   729: '-YB4 OP3_RESERVE_1', class Errors, trigger "DB_ALARM_OP3_M_3" bit 8
   730: '-YB4 OP3_RESERVE_2', class Errors, trigger "DB_ALARM_OP3_M_3" bit 9
   731: '-YB4 OP3_RESERVE_3', class Errors, trigger "DB_ALARM_OP3_M_3" bit 10
   732: '-YB4 OP3_RESERVE_4', class Errors, trigger "DB_ALARM_OP3_M_3" bit 11
   733: '-YB4 OP3_RESERVE_5', class Errors, trigger "DB_ALARM_OP3_M_3" bit 12
   734: '-YB4 OP3_RESERVE_6', class Errors, trigger "DB_ALARM_OP3_M_3" bit 13
   735: '-YB4 OP3_RESERVE_7', class Errors, trigger "DB_ALARM_OP3_M_3" bit 14
   736: '-YB4 OP3_RESERVE_8', class Errors, trigger "DB_ALARM_OP3_M_3" bit 15
   737: 'OP3_N0 -YB5 Nespecifikovaný režim motoru AUTOMAT/MANUAL', class Errors, trigger "DB_ALARM_OP3_M_4" bit 0
   738: 'OP3_N0 -YB5 Externí alarm err 1', class Errors, trigger "DB_ALARM_OP3_M_4" bit 1
   739: 'OP3_N0 -YB5 Externí alarm err 2', class Errors, trigger "DB_ALARM_OP3_M_4" bit 2
   740: 'OP3_N0 -YB5 Externí alarm err 3', class Errors, trigger "DB_ALARM_OP3_M_4" bit 3
   741: 'OP3_N0 -YB5 Motor nemá splněny podmínky pro opuštění pozice HOME', class Errors, trigger "DB_ALARM_OP3_M_4" bit 4
   742: 'OP3_N0 -YB5 Motor nemá splněny podmínky pro opuštění pozice WORK', class Errors, trigger "DB_ALARM_OP3_M_4" bit 5
   743: 'OP3_N0 -YB5 Motor nedojel do požadované pozice WORK', class Errors, trigger "DB_ALARM_OP3_M_4" bit 6
   744: 'OP3_N0 -YB5 Motor nedojel do požadované pozice HOME', class Errors, trigger "DB_ALARM_OP3_M_4" bit 7
   745: '-YB5 OP3_RESERVE_1', class Errors, trigger "DB_ALARM_OP3_M_4" bit 8
   746: '-YB5 OP3_RESERVE_2', class Errors, trigger "DB_ALARM_OP3_M_4" bit 9
   747: '-YB5 OP3_RESERVE_3', class Errors, trigger "DB_ALARM_OP3_M_4" bit 10
   748: '-YB5 OP3_RESERVE_4', class Errors, trigger "DB_ALARM_OP3_M_4" bit 11
   749: '-YB5 OP3_RESERVE_5', class Errors, trigger "DB_ALARM_OP3_M_4" bit 12
   750: '-YB5 OP3_RESERVE_6', class Errors, trigger "DB_ALARM_OP3_M_4" bit 13
   751: '-YB5 OP3_RESERVE_7', class Errors, trigger "DB_ALARM_OP3_M_4" bit 14
   752: '-YB5 OP3_RESERVE_8', class Errors, trigger "DB_ALARM_OP3_M_4" bit 15
   753: 'OP3_N0 -YB6 Nespecifikovaný režim motoru AUTOMAT/MANUAL', class Errors, trigger "DB_ALARM_OP3_M_5" bit 0
   754: 'OP3_N0 -YB6 Externí alarm err 1', class Errors, trigger "DB_ALARM_OP3_M_5" bit 1
   755: 'OP3_N0 -YB6 Externí alarm err 2', class Errors, trigger "DB_ALARM_OP3_M_5" bit 2
   756: 'OP3_N0 -YB6 Externí alarm err 3', class Errors, trigger "DB_ALARM_OP3_M_5" bit 3
   757: 'OP3_N0 -YB6 Motor nemá splněny podmínky pro opuštění pozice HOME', class Errors, trigger "DB_ALARM_OP3_M_5" bit 4
   758: 'OP3_N0 -YB6 Motor nemá splněny podmínky pro opuštění pozice WORK', class Errors, trigger "DB_ALARM_OP3_M_5" bit 5
   759: 'OP3_N0 -YB6 Motor nedojel do požadované pozice WORK', class Errors, trigger "DB_ALARM_OP3_M_5" bit 6
   760: 'OP3_N0 -YB6 Motor nedojel do požadované pozice HOME', class Errors, trigger "DB_ALARM_OP3_M_5" bit 7
   761: '-YB6 OP3_RESERVE_1', class Errors, trigger "DB_ALARM_OP3_M_5" bit 8
   762: '-YB6 OP3_RESERVE_2', class Errors, trigger "DB_ALARM_OP3_M_5" bit 9
   763: '-YB6 OP3_RESERVE_3', class Errors, trigger "DB_ALARM_OP3_M_5" bit 10
   764: '-YB6 OP3_RESERVE_4', class Errors, trigger "DB_ALARM_OP3_M_5" bit 11
   765: '-YB6 OP3_RESERVE_5', class Errors, trigger "DB_ALARM_OP3_M_5" bit 12
   766: '-YB6 OP3_RESERVE_6', class Errors, trigger "DB_ALARM_OP3_M_5" bit 13
   767: '-YB6 OP3_RESERVE_7', class Errors, trigger "DB_ALARM_OP3_M_5" bit 14
   768: '-YB6 OP3_RESERVE_8', class Errors, trigger "DB_ALARM_OP3_M_5" bit 15
   769: 'OP3_N0 -YB7 Nespecifikovaný režim motoru AUTOMAT/MANUAL', class Errors, trigger "DB_ALARM_OP3_M_6" bit 0
   770: 'OP3_N0 -YB7 Externí alarm err 1', class Errors, trigger "DB_ALARM_OP3_M_6" bit 1
   771: 'OP3_N0 -YB7 Externí alarm err 2', class Errors, trigger "DB_ALARM_OP3_M_6" bit 2
   772: 'OP3_N0 -YB7 Externí alarm err 3', class Errors, trigger "DB_ALARM_OP3_M_6" bit 3
   773: 'OP3_N0 -YB7 Motor nemá splněny podmínky pro opuštění pozice HOME', class Errors, trigger "DB_ALARM_OP3_M_6" bit 4
   774: 'OP3_N0 -YB7 Motor nemá splněny podmínky pro opuštění pozice WORK', class Errors, trigger "DB_ALARM_OP3_M_6" bit 5
   775: 'OP3_N0 -YB7 Motor nedojel do požadované pozice WORK', class Errors, trigger "DB_ALARM_OP3_M_6" bit 6
   776: 'OP3_N0 -YB7 Motor nedojel do požadované pozice HOME', class Errors, trigger "DB_ALARM_OP3_M_6" bit 7
   777: '-YB7 OP3_RESERVE_1', class Errors, trigger "DB_ALARM_OP3_M_6" bit 8
   778: '-YB7 OP3_RESERVE_2', class Errors, trigger "DB_ALARM_OP3_M_6" bit 9
   779: '-YB7 OP3_RESERVE_3', class Errors, trigger "DB_ALARM_OP3_M_6" bit 10
   780: '-YB7 OP3_RESERVE_4', class Errors, trigger "DB_ALARM_OP3_M_6" bit 11
   781: '-YB7 OP3_RESERVE_5', class Errors, trigger "DB_ALARM_OP3_M_6" bit 12
   782: '-YB7 OP3_RESERVE_6', class Errors, trigger "DB_ALARM_OP3_M_6" bit 13
   783: '-YB7 OP3_RESERVE_7', class Errors, trigger "DB_ALARM_OP3_M_6" bit 14
   784: '-YB7 OP3_RESERVE_8', class Errors, trigger "DB_ALARM_OP3_M_6" bit 15
   785: 'OP3_N0 -YB8 Nespecifikovaný režim motoru AUTOMAT/MANUAL', class Errors, trigger "DB_ALARM_OP3_M_7" bit 0
   786: 'OP3_N0 -YB8 Externí alarm err 1', class Errors, trigger "DB_ALARM_OP3_M_7" bit 1
   787: 'OP3_N0 -YB8 Externí alarm err 2', class Errors, trigger "DB_ALARM_OP3_M_7" bit 2
   788: 'OP3_N0 -YB8 Externí alarm err 3', class Errors, trigger "DB_ALARM_OP3_M_7" bit 3
   789: 'OP3_N0 -YB8 Motor nemá splněny podmínky pro opuštění pozice HOME', class Errors, trigger "DB_ALARM_OP3_M_7" bit 4
   790: 'OP3_N0 -YB8 Motor nemá splněny podmínky pro opuštění pozice WORK', class Errors, trigger "DB_ALARM_OP3_M_7" bit 5
   791: 'OP3_N0 -YB8 Motor nedojel do požadované pozice WORK', class Errors, trigger "DB_ALARM_OP3_M_7" bit 6
   792: 'OP3_N0 -YB8 Motor nedojel do požadované pozice HOME', class Errors, trigger "DB_ALARM_OP3_M_7" bit 7
   793: '-YB8 OP3_RESERVE_1', class Errors, trigger "DB_ALARM_OP3_M_7" bit 8
   794: '-YB8 OP3_RESERVE_2', class Errors, trigger "DB_ALARM_OP3_M_7" bit 9
   795: '-YB8 OP3_RESERVE_3', class Errors, trigger "DB_ALARM_OP3_M_7" bit 10
   796: '-YB8 OP3_RESERVE_4', class Errors, trigger "DB_ALARM_OP3_M_7" bit 11
   797: '-YB8 OP3_RESERVE_5', class Errors, trigger "DB_ALARM_OP3_M_7" bit 12
   798: '-YB8 OP3_RESERVE_6', class Errors, trigger "DB_ALARM_OP3_M_7" bit 13
   799: '-YB8 OP3_RESERVE_7', class Errors, trigger "DB_ALARM_OP3_M_7" bit 14
   800: '-YB8 OP3_RESERVE_8', class Errors, trigger "DB_ALARM_OP3_M_7" bit 15
   801: 'OP3_N0 Nespecifikovaný režim motoru AUTOMAT/MANUAL', class Errors, trigger "DB_ALARM_OP3_M_8" bit 0
   802: 'OP3_N0 Externí alarm err 1', class Errors, trigger "DB_ALARM_OP3_M_8" bit 1
   803: 'OP3_N0 Externí alarm err 2', class Errors, trigger "DB_ALARM_OP3_M_8" bit 2
   804: 'OP3_N0 Externí alarm err 3', class Errors, trigger "DB_ALARM_OP3_M_8" bit 3
   805: 'OP3_N0 Motor nemá splněny podmínky pro opuštění pozice HOME', class Errors, trigger "DB_ALARM_OP3_M_8" bit 4
   806: 'OP3_N0 Motor nemá splněny podmínky pro opuštění pozice WORK', class Errors, trigger "DB_ALARM_OP3_M_8" bit 5
   807: 'OP3_N0 Motor nedojel do požadované pozice WORK', class Errors, trigger "DB_ALARM_OP3_M_8" bit 6
   808: 'OP3_N0 Motor nedojel do požadované pozice HOME', class Errors, trigger "DB_ALARM_OP3_M_8" bit 7
   809: 'OP3_RESERVE_1', class Errors, trigger "DB_ALARM_OP3_M_8" bit 8
   810: 'OP3_RESERVE_2', class Errors, trigger "DB_ALARM_OP3_M_8" bit 9
   811: 'OP3_RESERVE_3', class Errors, trigger "DB_ALARM_OP3_M_8" bit 10
   812: 'OP3_RESERVE_4', class Errors, trigger "DB_ALARM_OP3_M_8" bit 11
   813: 'OP3_RESERVE_5', class Errors, trigger "DB_ALARM_OP3_M_8" bit 12
   814: 'OP3_RESERVE_6', class Errors, trigger "DB_ALARM_OP3_M_8" bit 13
   815: 'OP3_RESERVE_7', class Errors, trigger "DB_ALARM_OP3_M_8" bit 14
   816: 'OP3_RESERVE_8', class Errors, trigger "DB_ALARM_OP3_M_8" bit 15
   817: 'OP3_N0 Nespecifikovaný režim motoru AUTOMAT/MANUAL', class Errors, trigger "DB_ALARM_OP3_M_9" bit 0
   818: 'OP3_N0 Externí alarm err 1', class Errors, trigger "DB_ALARM_OP3_M_9" bit 1
   819: 'OP3_N0 Externí alarm err 2', class Errors, trigger "DB_ALARM_OP3_M_9" bit 2
   820: 'OP3_N0 Externí alarm err 3', class Errors, trigger "DB_ALARM_OP3_M_9" bit 3
   821: 'OP3_N0 Motor nemá splněny podmínky pro opuštění pozice HOME', class Errors, trigger "DB_ALARM_OP3_M_9" bit 4
   822: 'OP3_N0 Motor nemá splněny podmínky pro opuštění pozice WORK', class Errors, trigger "DB_ALARM_OP3_M_9" bit 5
   823: 'OP3_N0 Motor nedojel do požadované pozice WORK', class Errors, trigger "DB_ALARM_OP3_M_9" bit 6
   824: 'OP3_N0 Motor nedojel do požadované pozice HOME', class Errors, trigger "DB_ALARM_OP3_M_9" bit 7
   825: 'OP3_RESERVE_1', class Errors, trigger "DB_ALARM_OP3_M_9" bit 8
   826: 'OP3_RESERVE_2', class Errors, trigger "DB_ALARM_OP3_M_9" bit 9
   827: 'OP3_RESERVE_3', class Errors, trigger "DB_ALARM_OP3_M_9" bit 10
   828: 'OP3_RESERVE_4', class Errors, trigger "DB_ALARM_OP3_M_9" bit 11
   829: 'OP3_RESERVE_5', class Errors, trigger "DB_ALARM_OP3_M_9" bit 12
   830: 'OP3_RESERVE_6', class Errors, trigger "DB_ALARM_OP3_M_9" bit 13
   831: 'OP3_RESERVE_7', class Errors, trigger "DB_ALARM_OP3_M_9" bit 14
   832: 'OP3_RESERVE_8', class Errors, trigger "DB_ALARM_OP3_M_9" bit 15
   833: 'OP3_N0 Nespecifikovaný režim motoru AUTOMAT/MANUAL', class Errors, trigger "DB_ALARM_OP3_M_10" bit 0
   834: 'OP3_N0 Externí alarm err 1', class Errors, trigger "DB_ALARM_OP3_M_10" bit 1
   835: 'OP3_N0 Externí alarm err 2', class Errors, trigger "DB_ALARM_OP3_M_10" bit 2
   836: 'OP3_N0 Externí alarm err 3', class Errors, trigger "DB_ALARM_OP3_M_10" bit 3
   837: 'OP3_N0 Motor nemá splněny podmínky pro opuštění pozice HOME', class Errors, trigger "DB_ALARM_OP3_M_10" bit 4
   838: 'OP3_N0 Motor nemá splněny podmínky pro opuštění pozice WORK', class Errors, trigger "DB_ALARM_OP3_M_10" bit 5
   839: 'OP3_N0 Motor nedojel do požadované pozice WORK', class Errors, trigger "DB_ALARM_OP3_M_10" bit 6
   840: 'OP3_N0 Motor nedojel do požadované pozice HOME', class Errors, trigger "DB_ALARM_OP3_M_10" bit 7
   841: 'OP3_RESERVE_1', class Errors, trigger "DB_ALARM_OP3_M_10" bit 8
   842: 'OP3_RESERVE_2', class Errors, trigger "DB_ALARM_OP3_M_10" bit 9
   843: 'OP3_RESERVE_3', class Errors, trigger "DB_ALARM_OP3_M_10" bit 10
   844: 'OP3_RESERVE_4', class Errors, trigger "DB_ALARM_OP3_M_10" bit 11
   845: 'OP3_RESERVE_5', class Errors, trigger "DB_ALARM_OP3_M_10" bit 12
   846: 'OP3_RESERVE_6', class Errors, trigger "DB_ALARM_OP3_M_10" bit 13
   847: 'OP3_RESERVE_7', class Errors, trigger "DB_ALARM_OP3_M_10" bit 14
   848: 'OP3_RESERVE_8', class Errors, trigger "DB_ALARM_OP3_M_10" bit 15
   849: 'OP3_N0 Nespecifikovaný režim motoru AUTOMAT/MANUAL', class Errors, trigger "DB_ALARM_OP3_M_11" bit 0
   850: 'OP3_N0 Externí alarm err 1', class Errors, trigger "DB_ALARM_OP3_M_11" bit 1
   851: 'OP3_N0 Externí alarm err 2', class Errors, trigger "DB_ALARM_OP3_M_11" bit 2
   852: 'OP3_N0 Externí alarm err 3', class Errors, trigger "DB_ALARM_OP3_M_11" bit 3
   853: 'OP3_N0 Motor nemá splněny podmínky pro opuštění pozice HOME', class Errors, trigger "DB_ALARM_OP3_M_11" bit 4
   854: 'OP3_N0 Motor nemá splněny podmínky pro opuštění pozice WORK', class Errors, trigger "DB_ALARM_OP3_M_11" bit 5
   855: 'OP3_N0 Motor nedojel do požadované pozice WORK', class Errors, trigger "DB_ALARM_OP3_M_11" bit 6
   856: 'OP3_N0 Motor nedojel do požadované pozice HOME', class Errors, trigger "DB_ALARM_OP3_M_11" bit 7
   857: 'OP3_RESERVE_1', class Errors, trigger "DB_ALARM_OP3_M_11" bit 8
   858: 'OP3_RESERVE_2', class Errors, trigger "DB_ALARM_OP3_M_11" bit 9
   859: 'OP3_RESERVE_3', class Errors, trigger "DB_ALARM_OP3_M_11" bit 10
   860: 'OP3_RESERVE_4', class Errors, trigger "DB_ALARM_OP3_M_11" bit 11
   861: 'OP3_RESERVE_5', class Errors, trigger "DB_ALARM_OP3_M_11" bit 12
   862: 'OP3_RESERVE_6', class Errors, trigger "DB_ALARM_OP3_M_11" bit 13
   863: 'OP3_RESERVE_7', class Errors, trigger "DB_ALARM_OP3_M_11" bit 14
   864: 'OP3_RESERVE_8', class Errors, trigger "DB_ALARM_OP3_M_11" bit 15
   865: 'OP3_N0 Nespecifikovaný režim motoru AUTOMAT/MANUAL', class Errors, trigger "DB_ALARM_OP3_M_12" bit 0
   866: 'OP3_N0 Externí alarm err 1', class Errors, trigger "DB_ALARM_OP3_M_12" bit 1
   867: 'OP3_N0 Externí alarm err 2', class Errors, trigger "DB_ALARM_OP3_M_12" bit 2
   868: 'OP3_N0 Externí alarm err 3', class Errors, trigger "DB_ALARM_OP3_M_12" bit 3
   869: 'OP3_N0 Motor nemá splněny podmínky pro opuštění pozice HOME', class Errors, trigger "DB_ALARM_OP3_M_12" bit 4
   870: 'OP3_N0 Motor nemá splněny podmínky pro opuštění pozice WORK', class Errors, trigger "DB_ALARM_OP3_M_12" bit 5
   871: 'OP3_N0 Motor nedojel do požadované pozice WORK', class Errors, trigger "DB_ALARM_OP3_M_12" bit 6
   872: 'OP3_N0 Motor nedojel do požadované pozice HOME', class Errors, trigger "DB_ALARM_OP3_M_12" bit 7
   873: 'OP3_RESERVE_1', class Errors, trigger "DB_ALARM_OP3_M_12" bit 8
   874: 'OP3_RESERVE_2', class Errors, trigger "DB_ALARM_OP3_M_12" bit 9
   875: 'OP3_RESERVE_3', class Errors, trigger "DB_ALARM_OP3_M_12" bit 10
   876: 'OP3_RESERVE_4', class Errors, trigger "DB_ALARM_OP3_M_12" bit 11
   877: 'OP3_RESERVE_5', class Errors, trigger "DB_ALARM_OP3_M_12" bit 12
   878: 'OP3_RESERVE_6', class Errors, trigger "DB_ALARM_OP3_M_12" bit 13
   879: 'OP3_RESERVE_7', class Errors, trigger "DB_ALARM_OP3_M_12" bit 14
   880: 'OP3_RESERVE_8', class Errors, trigger "DB_ALARM_OP3_M_12" bit 15
   881: 'OP3_N0 Nespecifikovaný režim motoru AUTOMAT/MANUAL', class Errors, trigger "DB_ALARM_OP3_M_13" bit 0
   882: 'OP3_N0 Externí alarm err 1', class Errors, trigger "DB_ALARM_OP3_M_13" bit 1
   883: 'OP3_N0 Externí alarm err 2', class Errors, trigger "DB_ALARM_OP3_M_13" bit 2
   884: 'OP3_N0 Externí alarm err 3', class Errors, trigger "DB_ALARM_OP3_M_13" bit 3
   885: 'OP3_N0 Motor nemá splněny podmínky pro opuštění pozice HOME', class Errors, trigger "DB_ALARM_OP3_M_13" bit 4
   886: 'OP3_N0 Motor nemá splněny podmínky pro opuštění pozice WORK', class Errors, trigger "DB_ALARM_OP3_M_13" bit 5
   887: 'OP3_N0 Motor nedojel do požadované pozice WORK', class Errors, trigger "DB_ALARM_OP3_M_13" bit 6
   888: 'OP3_N0 Motor nedojel do požadované pozice HOME', class Errors, trigger "DB_ALARM_OP3_M_13" bit 7
   889: 'OP3_RESERVE_1', class Errors, trigger "DB_ALARM_OP3_M_13" bit 8
   890: 'OP3_RESERVE_2', class Errors, trigger "DB_ALARM_OP3_M_13" bit 9
   891: 'OP3_RESERVE_3', class Errors, trigger "DB_ALARM_OP3_M_13" bit 10
   892: 'OP3_RESERVE_4', class Errors, trigger "DB_ALARM_OP3_M_13" bit 11
   893: 'OP3_RESERVE_5', class Errors, trigger "DB_ALARM_OP3_M_13" bit 12
   894: 'OP3_RESERVE_6', class Errors, trigger "DB_ALARM_OP3_M_13" bit 13
   895: 'OP3_RESERVE_7', class Errors, trigger "DB_ALARM_OP3_M_13" bit 14
   896: 'OP3_RESERVE_8', class Errors, trigger "DB_ALARM_OP3_M_13" bit 15
   897: 'OP3_N0 Nespecifikovaný režim motoru AUTOMAT/MANUAL', class Errors, trigger "DB_ALARM_OP3_M_14" bit 0
   898: 'OP3_N0 Externí alarm err 1', class Errors, trigger "DB_ALARM_OP3_M_14" bit 1
   899: 'OP3_N0 Externí alarm err 2', class Errors, trigger "DB_ALARM_OP3_M_14" bit 2
   900: 'OP3_N0 Externí alarm err 3', class Errors, trigger "DB_ALARM_OP3_M_14" bit 3
   901: 'OP3_N0 Motor nemá splněny podmínky pro opuštění pozice HOME', class Errors, trigger "DB_ALARM_OP3_M_14" bit 4
   902: 'OP3_N0 Motor nemá splněny podmínky pro opuštění pozice WORK', class Errors, trigger "DB_ALARM_OP3_M_14" bit 5
   903: 'OP3_N0 Motor nedojel do požadované pozice WORK', class Errors, trigger "DB_ALARM_OP3_M_14" bit 6
   904: 'OP3_N0 Motor nedojel do požadované pozice HOME', class Errors, trigger "DB_ALARM_OP3_M_14" bit 7
   905: 'OP3_RESERVE_1', class Errors, trigger "DB_ALARM_OP3_M_14" bit 8
   906: 'OP3_RESERVE_2', class Errors, trigger "DB_ALARM_OP3_M_14" bit 9
   907: 'OP3_RESERVE_3', class Errors, trigger "DB_ALARM_OP3_M_14" bit 10
   908: 'OP3_RESERVE_4', class Errors, trigger "DB_ALARM_OP3_M_14" bit 11
   909: 'OP3_RESERVE_5', class Errors, trigger "DB_ALARM_OP3_M_14" bit 12
   910: 'OP3_RESERVE_6', class Errors, trigger "DB_ALARM_OP3_M_14" bit 13
   911: 'OP3_RESERVE_7', class Errors, trigger "DB_ALARM_OP3_M_14" bit 14
   912: 'OP3_RESERVE_8', class Errors, trigger "DB_ALARM_OP3_M_14" bit 15
   913: 'OP3_N0 Nespecifikovaný režim motoru AUTOMAT/MANUAL', class Errors, trigger "DB_ALARM_OP3_M_15" bit 0
   914: 'OP3_N0 Externí alarm err 1', class Errors, trigger "DB_ALARM_OP3_M_15" bit 1
   915: 'OP3_N0 Externí alarm err 2', class Errors, trigger "DB_ALARM_OP3_M_15" bit 2
   916: 'OP3_N0 Externí alarm err 3', class Errors, trigger "DB_ALARM_OP3_M_15" bit 3
   917: 'OP3_N0 Motor nemá splněny podmínky pro opuštění pozice HOME', class Errors, trigger "DB_ALARM_OP3_M_15" bit 4
   918: 'OP3_N0 Motor nemá splněny podmínky pro opuštění pozice WORK', class Errors, trigger "DB_ALARM_OP3_M_15" bit 5
   919: 'OP3_N0 Motor nedojel do požadované pozice WORK', class Errors, trigger "DB_ALARM_OP3_M_15" bit 6
   920: 'OP3_N0 Motor nedojel do požadované pozice HOME', class Errors, trigger "DB_ALARM_OP3_M_15" bit 7
   921: 'OP3_RESERVE_1', class Errors, trigger "DB_ALARM_OP3_M_15" bit 8
   922: 'OP3_RESERVE_2', class Errors, trigger "DB_ALARM_OP3_M_15" bit 9
   923: 'OP3_RESERVE_3', class Errors, trigger "DB_ALARM_OP3_M_15" bit 10
   924: 'OP3_RESERVE_4', class Errors, trigger "DB_ALARM_OP3_M_15" bit 11
   925: 'OP3_RESERVE_5', class Errors, trigger "DB_ALARM_OP3_M_15" bit 12
   926: 'OP3_RESERVE_6', class Errors, trigger "DB_ALARM_OP3_M_15" bit 13
   927: 'OP3_RESERVE_7', class Errors, trigger "DB_ALARM_OP3_M_15" bit 14
   928: 'OP3_RESERVE_8', class Errors, trigger "DB_ALARM_OP3_M_15" bit 15
   129: 'Odsávací zařízení nereaguje. Otevřete dveře a zkontrolujte jej.', class Errors bit 0
   130: 'op_4_alrm_10', class Errors bit 0
   131: 'op_4_alrm_11', class Errors bit 0
   132: 'op_4_alrm_12', class Errors bit 0
   133: 'op_4_alrm_13', class Errors bit 0
   134: 'op_4_alrm_14', class Errors bit 0
   135: 'op_4_alrm_15', class Errors bit 0
   136: 'Odsávací zařízení nereaguje. Otevřete dveře a zkontrolujte jej.', class Errors bit 0
   137: 'op_4_alrm_2', class Errors bit 0
   138: 'op_4_alrm_3', class Errors bit 0
   139: 'op_4_alrm_4', class Errors bit 0
   140: 'op_4_alrm_5', class Errors bit 0
   141: 'op_4_alrm_6', class Errors bit 0
   142: 'op_4_alrm_7', class Errors bit 0
   143: 'op_4_alrm_8', class Errors bit 0
   144: 'OTEVŘEN BEZPEČNOSTNÍ KRYT (dveře 1)', class Errors bit 0
   929: 'op_4_N0 -Y7 Nespecifikovaný režim motoru AUTOMAT/MANUAL', class Errors bit 0
   930: 'op_4_N0 -Y7 Externí alarm err 1', class Errors bit 1
   931: 'op_4_-Y7 RESERVE_3', class Errors bit 10
   932: 'op_4_-Y7 RESERVE_4', class Errors bit 11
   933: 'op_4_-Y7 RESERVE_5', class Errors bit 12
   934: 'op_4_-Y7 RESERVE_6', class Errors bit 13
   935: 'op_4_-Y7 RESERVE_7', class Errors bit 14
   936: 'op_4_-Y7 RESERVE_8', class Errors bit 15
   937: 'op_4_N0 -Y7 Externí alarm err 2', class Errors bit 2
   938: 'op_4_N0 -Y7 Externí alarm err 3', class Errors bit 3
   939: 'op_4_N0 -Y7 Motor nemá splněny podmínky pro opuštění pozice HOME', class Errors bit 4
   940: 'op_4_N0 -Y7 Motor nemá splněny podmínky pro opuštění pozice WORK', class Errors bit 5
   941: 'op_4_N0 -Y7 Motor nedojel do požadované pozice WORK', class Errors bit 6
   942: 'op_4_N0 -Y7 Motor nedojel do požadované pozice HOME', class Errors bit 7
   943: 'op_4_-Y7 RESERVE_1', class Errors bit 8
   944: 'op_4_-Y7 RESERVE_2', class Errors bit 9
   945: 'op_4_N0 -Y9 Nespecifikovaný režim motoru AUTOMAT/MANUAL', class Errors bit 0
   946: 'op_4_N0 -Y9 Externí alarm err 1', class Errors bit 1
   947: 'op_4_RESERVE_3 -Y9', class Errors bit 10
   948: 'op_4_RESERVE_4 -Y9', class Errors bit 11
   949: 'op_4_RESERVE_5 -Y9', class Errors bit 12
   950: 'op_4_RESERVE_6 -Y9', class Errors bit 13
   951: 'op_4_RESERVE_7 -Y9', class Errors bit 14
   952: 'op_4_RESERVE_8 -Y9', class Errors bit 15
   953: 'op_4_N0 -Y9 Externí alarm err 2', class Errors bit 2
   954: 'op_4_N0 -Y9 Externí alarm err 3', class Errors bit 3
   955: 'op_4_N0 -Y9 Motor nemá splněny podmínky pro opuštění pozice HOME', class Errors bit 4
   956: 'op_4_N0 -Y9 Motor nemá splněny podmínky pro opuštění pozice WORK', class Errors bit 5
   957: 'op_4_N0 -Y9 Motor nedojel do požadované pozice WORK', class Errors bit 6
   958: 'op_4_N0 -Y9 Motor nedojel do požadované pozice HOME', class Errors bit 7
   959: 'op_4_RESERVE_1 -Y9', class Errors bit 8
   960: 'op_4_RESERVE_2 -Y9', class Errors bit 9
   961: 'op_4_N0 Nespecifikovaný režim motoru AUTOMAT/MANUAL', class Errors bit 0
   962: 'op_4_N0 Externí alarm err 1', class Errors bit 1
   963: 'op_4_RESERVE_3', class Errors bit 10
   964: 'op_4_RESERVE_4', class Errors bit 11
   965: 'op_4_RESERVE_5', class Errors bit 12
   966: 'op_4_RESERVE_6', class Errors bit 13
   967: 'op_4_RESERVE_7', class Errors bit 14
   968: 'op_4_RESERVE_8', class Errors bit 15
   969: 'op_4_N0 Externí alarm err 2', class Errors bit 2
   970: 'op_4_N0 Externí alarm err 3', class Errors bit 3
   971: 'op_4_N0 Motor nemá splněny podmínky pro opuštění pozice HOME', class Errors bit 4
   972: 'op_4_N0 Motor nemá splněny podmínky pro opuštění pozice WORK', class Errors bit 5
   973: 'op_4_N0 Motor nedojel do požadované pozice WORK', class Errors bit 6
   974: 'op_4_N0 Motor nedojel do požadované pozice HOME', class Errors bit 7
   975: 'op_4_RESERVE_1', class Errors bit 8
   976: 'op_4_RESERVE_2', class Errors bit 9
   977: 'op_4_N0 Nespecifikovaný režim motoru AUTOMAT/MANUAL', class Errors bit 0
   978: 'op_4_N0 Externí alarm err 1', class Errors bit 1
   979: 'op_4_RESERVE_3', class Errors bit 10
   980: 'op_4_RESERVE_4', class Errors bit 11
   981: 'op_4_RESERVE_5', class Errors bit 12
   982: 'op_4_RESERVE_6', class Errors bit 13
   983: 'op_4_RESERVE_7', class Errors bit 14
   984: 'op_4_RESERVE_8', class Errors bit 15
   985: 'op_4_N0 Externí alarm err 2', class Errors bit 2
   986: 'op_4_N0 Externí alarm err 3', class Errors bit 3
   987: 'op_4_N0 Motor nemá splněny podmínky pro opuštění pozice HOME', class Errors bit 4
   988: 'op_4_N0 Motor nemá splněny podmínky pro opuštění pozice WORK', class Errors bit 5
   989: 'op_4_N0 Motor nedojel do požadované pozice WORK', class Errors bit 6
   990: 'op_4_N0 Motor nedojel do požadované pozice HOME', class Errors bit 7
   991: 'op_4_RESERVE_1', class Errors bit 8
   992: 'op_4_RESERVE_2', class Errors bit 9
   993: 'op_4_N0 Nespecifikovaný režim motoru AUTOMAT/MANUAL', class Errors bit 0
   994: 'op_4_N0 Externí alarm err 1', class Errors bit 1
   995: 'op_4_RESERVE_3', class Errors bit 10
   996: 'op_4_RESERVE_4', class Errors bit 11
   997: 'op_4_RESERVE_5', class Errors bit 12
   998: 'op_4_RESERVE_6', class Errors bit 13
   999: 'op_4_RESERVE_7', class Errors bit 14
   1000: 'op_4_RESERVE_8', class Errors bit 15
   1001: 'op_4_N0 Externí alarm err 2', class Errors bit 2
   1002: 'op_4_N0 Externí alarm err 3', class Errors bit 3
   1003: 'op_4_N0 Motor nemá splněny podmínky pro opuštění pozice HOME', class Errors bit 4
   1004: 'op_4_N0 Motor nemá splněny podmínky pro opuštění pozice WORK', class Errors bit 5
   1005: 'op_4_N0 Motor nedojel do požadované pozice WORK', class Errors bit 6
   1006: 'op_4_N0 Motor nedojel do požadované pozice HOME', class Errors bit 7
   1007: 'op_4_RESERVE_1', class Errors bit 8
   1008: 'op_4_RESERVE_2', class Errors bit 9
   1009: 'op_4_N0 Nespecifikovaný režim motoru AUTOMAT/MANUAL', class Errors bit 0
   1010: 'op_4_N0 Externí alarm err 1', class Errors bit 1
   1011: 'op_4_RESERVE_3', class Errors bit 10
   1012: 'op_4_RESERVE_4', class Errors bit 11
   1013: 'op_4_RESERVE_5', class Errors bit 12
   1014: 'op_4_RESERVE_6', class Errors bit 13
   1015: 'op_4_RESERVE_7', class Errors bit 14
   1016: 'op_4_RESERVE_8', class Errors bit 15
   1017: 'op_4_N0 Externí alarm err 2', class Errors bit 2
   1018: 'op_4_N0 Externí alarm err 3', class Errors bit 3
   1019: 'op_4_N0 Motor nemá splněny podmínky pro opuštění pozice HOME', class Errors bit 4
   1020: 'op_4_N0 Motor nemá splněny podmínky pro opuštění pozice WORK', class Errors bit 5
   1021: 'op_4_N0 Motor nedojel do požadované pozice WORK', class Errors bit 6
   1022: 'op_4_N0 Motor nedojel do požadované pozice HOME', class Errors bit 7
   1023: 'op_4_RESERVE_1', class Errors bit 8
   1024: 'op_4_RESERVE_2', class Errors bit 9
   1025: 'op_4_N0 Nespecifikovaný režim motoru AUTOMAT/MANUAL', class Errors bit 0
   1026: 'op_4_N0 Externí alarm err 1', class Errors bit 1
   1027: 'op_4_RESERVE_3', class Errors bit 10
   1028: 'op_4_RESERVE_4', class Errors bit 11
   1029: 'op_4_RESERVE_5', class Errors bit 12
   1030: 'op_4_RESERVE_6', class Errors bit 13
   1031: 'op_4_RESERVE_7', class Errors bit 14
   1032: 'op_4_RESERVE_8', class Errors bit 15
   1033: 'op_4_N0 Externí alarm err 2', class Errors bit 2
   1034: 'op_4_N0 Externí alarm err 3', class Errors bit 3
   1035: 'op_4_N0 Motor nemá splněny podmínky pro opuštění pozice HOME', class Errors bit 4
   1036: 'op_4_N0 Motor nemá splněny podmínky pro opuštění pozice WORK', class Errors bit 5
   1037: 'op_4_N0 Motor nedojel do požadované pozice WORK', class Errors bit 6
   1038: 'op_4_N0 Motor nedojel do požadované pozice HOME', class Errors bit 7
   1039: 'op_4_RESERVE_1', class Errors bit 8
   1040: 'op_4_RESERVE_2', class Errors bit 9
   1041: 'op_4_N0 Nespecifikovaný režim motoru AUTOMAT/MANUAL', class Errors bit 0
   1042: 'op_4_N0 Externí alarm err 1', class Errors bit 1
   1043: 'op_4_RESERVE_3', class Errors bit 10
   1044: 'op_4_RESERVE_4', class Errors bit 11
   1045: 'op_4_RESERVE_5', class Errors bit 12
   1046: 'op_4_RESERVE_6', class Errors bit 13
   1047: 'op_4_RESERVE_7', class Errors bit 14
   1048: 'op_4_RESERVE_8', class Errors bit 15
   1049: 'op_4_N0 Externí alarm err 2', class Errors bit 2
   1050: 'op_4_N0 Externí alarm err 3', class Errors bit 3
   1051: 'op_4_N0 Motor nemá splněny podmínky pro opuštění pozice HOME', class Errors bit 4
   1052: 'op_4_N0 Motor nemá splněny podmínky pro opuštění pozice WORK', class Errors bit 5
   1053: 'op_4_N0 Motor nedojel do požadované pozice WORK', class Errors bit 6
   1054: 'op_4_N0 Motor nedojel do požadované pozice HOME', class Errors bit 7
   1055: 'op_4_RESERVE_1', class Errors bit 8
   1056: 'op_4_RESERVE_2', class Errors bit 9
   1057: 'op_4_N0 Nespecifikovaný režim motoru AUTOMAT/MANUAL', class Errors bit 0
   1058: 'op_4_N0 Externí alarm err 1', class Errors bit 1
   1059: 'op_4_RESERVE_3', class Errors bit 10
   1060: 'op_4_RESERVE_4', class Errors bit 11
   1061: 'op_4_RESERVE_5', class Errors bit 12
   1062: 'op_4_RESERVE_6', class Errors bit 13
   1063: 'op_4_RESERVE_7', class Errors bit 14
   1064: 'op_4_RESERVE_8', class Errors bit 15
   1065: 'op_4_N0 Externí alarm err 2', class Errors bit 2
   1066: 'op_4_N0 Externí alarm err 3', class Errors bit 3
   1067: 'op_4_N0 Motor nemá splněny podmínky pro opuštění pozice HOME', class Errors bit 4
   1068: 'op_4_N0 Motor nemá splněny podmínky pro opuštění pozice WORK', class Errors bit 5
   1069: 'op_4_N0 Motor nedojel do požadované pozice WORK', class Errors bit 6
   1070: 'op_4_N0 Motor nedojel do požadované pozice HOME', class Errors bit 7
   1071: 'op_4_RESERVE_1', class Errors bit 8
   1072: 'op_4_RESERVE_2', class Errors bit 9
   1073: 'op_4_N0 Nespecifikovaný režim motoru AUTOMAT/MANUAL', class Errors bit 0
   1074: 'op_4_N0 Externí alarm err 1', class Errors bit 1
   1075: 'op_4_RESERVE_3', class Errors bit 10
   1076: 'op_4_RESERVE_4', class Errors bit 11
   1077: 'op_4_RESERVE_5', class Errors bit 12
   1078: 'op_4_RESERVE_6', class Errors bit 13
   1079: 'op_4_RESERVE_7', class Errors bit 14
   1080: 'op_4_RESERVE_8', class Errors bit 15
   1081: 'op_4_N0 Externí alarm err 2', class Errors bit 2
   1082: 'op_4_N0 Externí alarm err 3', class Errors bit 3
   1083: 'op_4_N0 Motor nemá splněny podmínky pro opuštění pozice HOME', class Errors bit 4
   1084: 'op_4_N0 Motor nemá splněny podmínky pro opuštění pozice WORK', class Errors bit 5
   1085: 'op_4_N0 Motor nedojel do požadované pozice WORK', class Errors bit 6
   1086: 'op_4_N0 Motor nedojel do požadované pozice HOME', class Errors bit 7
   1087: 'op_4_RESERVE_1', class Errors bit 8
   1088: 'op_4_RESERVE_2', class Errors bit 9
   1089: 'op_4_N0 Nespecifikovaný režim motoru AUTOMAT/MANUAL', class Errors bit 0
   1090: 'op_4_N0 Externí alarm err 1', class Errors bit 1
   1091: 'op_4_RESERVE_3', class Errors bit 10
   1092: 'op_4_RESERVE_4', class Errors bit 11
   1093: 'op_4_RESERVE_5', class Errors bit 12
   1094: 'op_4_RESERVE_6', class Errors bit 13
   1095: 'op_4_RESERVE_7', class Errors bit 14
   1096: 'op_4_RESERVE_8', class Errors bit 15
   1097: 'op_4_N0 Externí alarm err 2', class Errors bit 2
   1098: 'op_4_N0 Externí alarm err 3', class Errors bit 3
   1099: 'op_4_N0 Motor nemá splněny podmínky pro opuštění pozice HOME', class Errors bit 4
   1100: 'op_4_N0 Motor nemá splněny podmínky pro opuštění pozice WORK', class Errors bit 5
   1101: 'op_4_N0 Motor nedojel do požadované pozice WORK', class Errors bit 6
   1102: 'op_4_N0 Motor nedojel do požadované pozice HOME', class Errors bit 7
   1103: 'op_4_RESERVE_1', class Errors bit 8
   1104: 'op_4_RESERVE_2', class Errors bit 9
   1105: 'op_4_N0 Nespecifikovaný režim motoru AUTOMAT/MANUAL', class Errors bit 0
   1106: 'op_4_N0 Externí alarm err 1', class Errors bit 1
   1107: 'op_4_RESERVE_3', class Errors bit 10
   1108: 'op_4_RESERVE_4', class Errors bit 11
   1109: 'op_4_RESERVE_5', class Errors bit 12
   1110: 'op_4_RESERVE_6', class Errors bit 13
   1111: 'op_4_RESERVE_7', class Errors bit 14
   1112: 'op_4_RESERVE_8', class Errors bit 15
   1113: 'op_4_N0 Externí alarm err 2', class Errors bit 2
   1114: 'op_4_N0 Externí alarm err 3', class Errors bit 3
   1115: 'op_4_N0 Motor nemá splněny podmínky pro opuštění pozice HOME', class Errors bit 4
   1116: 'op_4_N0 Motor nemá splněny podmínky pro opuštění pozice WORK', class Errors bit 5
   1117: 'op_4_N0 Motor nedojel do požadované pozice WORK', class Errors bit 6
   1118: 'op_4_N0 Motor nedojel do požadované pozice HOME', class Errors bit 7
   1119: 'op_4_RESERVE_1', class Errors bit 8
   1120: 'op_4_RESERVE_2', class Errors bit 9
   1121: 'op_4_N0 Nespecifikovaný režim motoru AUTOMAT/MANUAL', class Errors bit 0
   1122: 'op_4_N0 Externí alarm err 1', class Errors bit 1
   1123: 'op_4_RESERVE_3', class Errors bit 10
   1124: 'op_4_RESERVE_4', class Errors bit 11
   1125: 'op_4_RESERVE_5', class Errors bit 12
   1126: 'op_4_RESERVE_6', class Errors bit 13
   1127: 'op_4_RESERVE_7', class Errors bit 14
   1128: 'op_4_RESERVE_8', class Errors bit 15
   1129: 'op_4_N0 Externí alarm err 2', class Errors bit 2
   1130: 'op_4_N0 Externí alarm err 3', class Errors bit 3
   1131: 'op_4_N0 Motor nemá splněny podmínky pro opuštění pozice HOME', class Errors bit 4
   1132: 'op_4_N0 Motor nemá splněny podmínky pro opuštění pozice WORK', class Errors bit 5
   1133: 'op_4_N0 Motor nedojel do požadované pozice WORK', class Errors bit 6
   1134: 'op_4_N0 Motor nedojel do požadované pozice HOME', class Errors bit 7
   1135: 'op_4_RESERVE_1', class Errors bit 8
   1136: 'op_4_RESERVE_2', class Errors bit 9
   1137: 'op_4_N0 Nespecifikovaný režim motoru AUTOMAT/MANUAL', class Errors bit 0
   1138: 'op_4_N0 Externí alarm err 1', class Errors bit 1
   1139: 'op_4_RESERVE_3', class Errors bit 10
   1140: 'op_4_RESERVE_4', class Errors bit 11
   1141: 'op_4_RESERVE_5', class Errors bit 12
   1142: 'op_4_RESERVE_6', class Errors bit 13
   1143: 'op_4_RESERVE_7', class Errors bit 14
   1144: 'op_4_RESERVE_8', class Errors bit 15
   1145: 'op_4_N0 Externí alarm err 2', class Errors bit 2
   1146: 'op_4_N0 Externí alarm err 3', class Errors bit 3
   1147: 'op_4_N0 Motor nemá splněny podmínky pro opuštění pozice HOME', class Errors bit 4
   1148: 'op_4_N0 Motor nemá splněny podmínky pro opuštění pozice WORK', class Errors bit 5
   1149: 'op_4_N0 Motor nedojel do požadované pozice WORK', class Errors bit 6
   1150: 'op_4_N0 Motor nedojel do požadované pozice HOME', class Errors bit 7
   1151: 'op_4_RESERVE_1', class Errors bit 8
   1152: 'op_4_RESERVE_2', class Errors bit 9
   1153: 'op_4_N0 Nespecifikovaný režim motoru AUTOMAT/MANUAL', class Errors bit 0
   1154: 'op_4_N0 Externí alarm err 1', class Errors bit 1
   1155: 'op_4_RESERVE_3', class Errors bit 10
   1156: 'op_4_RESERVE_4', class Errors bit 11
   1157: 'op_4_RESERVE_5', class Errors bit 12
   1158: 'op_4_RESERVE_6', class Errors bit 13
   1159: 'op_4_RESERVE_7', class Errors bit 14
   1160: 'op_4_RESERVE_8', class Errors bit 15
   1161: 'op_4_N0 Externí alarm err 2', class Errors bit 2
   1162: 'op_4_N0 Externí alarm err 3', class Errors bit 3
   1163: 'op_4_N0 Motor nemá splněny podmínky pro opuštění pozice HOME', class Errors bit 4
   1164: 'op_4_N0 Motor nemá splněny podmínky pro opuštění pozice WORK', class Errors bit 5
   1165: 'op_4_N0 Motor nedojel do požadované pozice WORK', class Errors bit 6
   1166: 'op_4_N0 Motor nedojel do požadované pozice HOME', class Errors bit 7
   1167: 'op_4_RESERVE_1', class Errors bit 8
   1168: 'op_4_RESERVE_2', class Errors bit 9
   1169: 'op_4_N0 Nespecifikovaný režim motoru AUTOMAT/MANUAL', class Errors bit 0
   1170: 'op_4_N0 Externí alarm err 1', class Errors bit 1
   1171: 'op_4_RESERVE_3', class Errors bit 10
   1172: 'op_4_RESERVE_4', class Errors bit 11
   1173: 'op_4_RESERVE_5', class Errors bit 12
   1174: 'op_4_RESERVE_6', class Errors bit 13
   1175: 'op_4_RESERVE_7', class Errors bit 14
   1176: 'op_4_RESERVE_8', class Errors bit 15
   1177: 'op_4_N0 Externí alarm err 2', class Errors bit 2
   1178: 'op_4_N0 Externí alarm err 3', class Errors bit 3
   1179: 'op_4_N0 Motor nemá splněny podmínky pro opuštění pozice HOME', class Errors bit 4
   1180: 'op_4_N0 Motor nemá splněny podmínky pro opuštění pozice WORK', class Errors bit 5
   1181: 'op_4_N0 Motor nedojel do požadované pozice WORK', class Errors bit 6
   1182: 'op_4_N0 Motor nedojel do požadované pozice HOME', class Errors bit 7
   1183: 'op_4_RESERVE_1', class Errors bit 8
   1184: 'op_4_RESERVE_2', class Errors bit 9
   1185: 'op_4_wrong_1', class warning_individual bit 0
   1186: 'op_4_wrong_10', class warning_individual bit 9
   1187: 'op_4_wrong_11', class warning_individual bit 10
   1188: 'op_4_wrong_12', class warning_individual bit 11
   1189: 'op_4_wrong_13', class warning_individual bit 12
   1190: 'op_4_wrong_14', class warning_individual bit 13
   1191: 'op_4_wrong_15', class warning_individual bit 14
   1192: 'op_4_wrong_16', class warning_individual bit 15
   1193: 'op_4_wrong_2', class warning_individual bit 1
   1194: 'op_4_wrong_3', class warning_individual bit 2
   1195: 'op_4_wrong_4', class warning_individual bit 3
   1196: 'op_4_wrong_5', class warning_individual bit 4
   1197: 'op_4_wrong_6', class warning_individual bit 5
   1198: 'op_4_wrong_7', class warning_individual bit 6
   1199: 'op_4_wrong_8', class warning_individual bit 7
   1200: 'op_4_wrong_9', class warning_individual bit 8
   1201: 'op_2_wrong_12', class warning_individual, trigger "DB_ALARM_wrong_op_2" bit 11
   1202: 'op_2_wrong_11', class warning_individual, trigger "DB_ALARM_wrong_op_2" bit 10
   1203: 'op_2_wrong_10', class warning_individual, trigger "DB_ALARM_wrong_op_2" bit 9
   1204: 'op_2_wrong_9', class warning_individual, trigger "DB_ALARM_wrong_op_2" bit 8
   1205: 'op_2_wrong_8', class warning_individual, trigger "DB_ALARM_wrong_op_2" bit 7
   1206: 'op_2_wrong_6', class warning_individual, trigger "DB_ALARM_wrong_op_2" bit 5
   1207: 'op_2_wrong_5', class warning_individual, trigger "DB_ALARM_wrong_op_2" bit 4
   1208: 'op_2_wrong_4', class warning_individual, trigger "DB_ALARM_wrong_op_2" bit 3
   1209: 'op_2_wrong_3', class warning_individual, trigger "DB_ALARM_wrong_op_2" bit 2
   1210: 'op_2_wrong_2', class warning_individual, trigger "DB_ALARM_wrong_op_2" bit 1
   1211: 'op_2_wrong_1', class warning_individual, trigger "DB_ALARM_wrong_op_2" bit 0
   1212: 'op_3_wrong_14', class warning_individual, trigger "DB_ALARM_wrong_op_3" bit 13
   1213: 'op_2_wrong_7', class warning_individual, trigger "DB_ALARM_wrong_op_2" bit 6
   1214: 'op_1_wrong_15', class warning_individual, trigger "DB_ALARM_wrong_op_1" bit 14
   1215: 'op_2_wrong_13', class warning_individual, trigger "DB_ALARM_wrong_op_2" bit 12
   1216: 'op_2_wrong_15', class warning_individual, trigger "DB_ALARM_wrong_op_2" bit 14
   1217: 'op_2_wrong_16', class warning_individual, trigger "DB_ALARM_wrong_op_2" bit 15
   1218: 'op_3_wrong_13', class warning_individual, trigger "DB_ALARM_wrong_op_3" bit 12
   1219: 'op_3_wrong_12', class warning_individual, trigger "DB_ALARM_wrong_op_3" bit 11
   1220: 'op_3_wrong_1', class warning_individual, trigger "DB_ALARM_wrong_op_3" bit 0
   1221: 'op_3_wrong_2', class warning_individual, trigger "DB_ALARM_wrong_op_3" bit 1
   1222: 'op_3_wrong_3', class warning_individual, trigger "DB_ALARM_wrong_op_3" bit 2
   1223: 'op_3_wrong_4', class warning_individual, trigger "DB_ALARM_wrong_op_3" bit 3
   1224: 'op_3_wrong_5', class warning_individual, trigger "DB_ALARM_wrong_op_3" bit 4
   1225: 'op_3_wrong_6', class warning_individual, trigger "DB_ALARM_wrong_op_3" bit 5
   1226: 'op_3_wrong_7', class warning_individual, trigger "DB_ALARM_wrong_op_3" bit 6
   1227: 'op_3_wrong_8', class warning_individual, trigger "DB_ALARM_wrong_op_3" bit 7
   1228: 'op_3_wrong_9', class warning_individual, trigger "DB_ALARM_wrong_op_3" bit 8
   1229: 'op_2_wrong_14', class warning_individual, trigger "DB_ALARM_wrong_op_2" bit 13
   1230: 'op_1_wrong_16', class warning_individual, trigger "DB_ALARM_wrong_op_1" bit 15
   1231: 'op_3_wrong_11', class warning_individual, trigger "DB_ALARM_wrong_op_3" bit 10
   1232: 'op_1_wrong_14', class warning_individual, trigger "DB_ALARM_wrong_op_1" bit 13
   1233: 'wrong_line_1', class warning_individual, trigger "DB_ALARM_wrong_line" bit 0
   1234: 'wrong_line_2', class warning_individual, trigger "DB_ALARM_wrong_line" bit 1
   1235: 'wrong_line_3', class warning_individual, trigger "DB_ALARM_wrong_line" bit 2
   1236: 'wrong_line_4', class warning_individual, trigger "DB_ALARM_wrong_line" bit 3
   1237: 'wrong_line_5', class warning_individual, trigger "DB_ALARM_wrong_line" bit 4
   1238: 'wrong_line_6', class warning_individual, trigger "DB_ALARM_wrong_line" bit 5
   1239: 'Čelisti ropex je nutné zkontrolovat', class warning_individual, trigger "DB_ALARM_wrong_line" bit 6
   1240: 'Ropex autocal aktivní', class warning_individual, trigger "DB_ALARM_wrong_line" bit 7
   1241: 'Běží inicializace VYČKEJTE', class warning_individual, trigger "DB_ALARM_wrong_line" bit 8
   1242: 'Globální upozornění - zařízení nebo část není ve standardu', class warning_individual, trigger "DB_ALARM_wrong_line" bit 9
   1243: 'wrong_line_11', class warning_individual, trigger "DB_ALARM_wrong_line" bit 10
   1244: 'wrong_line_12', class warning_individual, trigger "DB_ALARM_wrong_line" bit 11
   1245: 'wrong_line_13', class warning_individual, trigger "DB_ALARM_wrong_line" bit 12
   1246: 'wrong_line_14', class warning_individual, trigger "DB_ALARM_wrong_line" bit 13
   1247: 'Zařízení ropex není ve standartním stavu otevřete obrazovku ROPEX + PODÉLNÉ ČELISTI a zkontorlujte hlášení', class warning_individual, trigger "DB_ALARM_wrong_line" bit 14
   1248: 'Ropex provádí kalibraci vyčkejte (ROPEX + PODÉLNÉ ČELISTI)', class warning_individual, trigger "DB_ALARM_wrong_line" bit 15
   1249: 'op_3_wrong_16', class warning_individual, trigger "DB_ALARM_wrong_op_3" bit 15
   1250: 'op_1_wrong_13', class warning_individual, trigger "DB_ALARM_wrong_op_1" bit 12
   1251: 'op_1_wrong_12', class warning_individual, trigger "DB_ALARM_wrong_op_1" bit 11
   1252: 'op_1_wrong_11', class warning_individual, trigger "DB_ALARM_wrong_op_1" bit 10
   1253: 'op_1_wrong_10', class warning_individual, trigger "DB_ALARM_wrong_op_1" bit 9
   1254: 'op_1_wrong_9', class warning_individual, trigger "DB_ALARM_wrong_op_1" bit 8
   1255: 'op_1_wrong_8', class warning_individual, trigger "DB_ALARM_wrong_op_1" bit 7
   1256: 'op_3_wrong_10', class warning_individual, trigger "DB_ALARM_wrong_op_3" bit 9
   1257: 'op_1_wrong_7', class warning_individual, trigger "DB_ALARM_wrong_op_1" bit 6
   1258: 'op_1_wrong_5', class warning_individual, trigger "DB_ALARM_wrong_op_1" bit 4
   1259: 'op_1_wrong_4', class warning_individual, trigger "DB_ALARM_wrong_op_1" bit 3
   1260: 'op_1_wrong_3', class warning_individual, trigger "DB_ALARM_wrong_op_1" bit 2
   1261: 'op_1_wrong_2', class warning_individual, trigger "DB_ALARM_wrong_op_1" bit 1
   1262: 'op_1_wrong_1', class warning_individual, trigger "DB_ALARM_wrong_op_1" bit 0
   1263: 'op_3_wrong_15', class warning_individual, trigger "DB_ALARM_wrong_op_3" bit 14
   1264: 'op_1_wrong_6', class warning_individual, trigger "DB_ALARM_wrong_op_1" bit 5
   1265: 'DOŠLA FOLIE -21B3', class Errors, trigger "DB_ALARM_alarm_op_2" bit 6
   1266: 'op_3_alarm_1', class Errors, trigger "DB_ALARM_alarm_op_3" bit 0
   1267: 'op_4_alrm_2', class Errors, trigger "DB_ALARM_alarm_op_4" bit 8
   1268: 'op_4_alrm_3', class Errors, trigger "DB_ALARM_alarm_op_4" bit 9
   1269: 'SERVO SELHÁNÍ BLOKU OVLÁDÁNÍ "POWER" (KONTAKTUJTE LIFTEC)', class Errors, trigger "DB_ALARM_alarm_op_2" bit 15
   1270: 'ROPEX ALARM ZKONTROLUJTE OBRAZOVKU (ROPEX + PODÉLNÉ ČELISTI)', class Errors, trigger "DB_ALARM_alarm_op_2" bit 14
   1271: 'PORUCHA ROPEXU PROVEĎTE INICIALIZACI ( PŘEPNUTÍM REŽIMŮ)', class Errors, trigger "DB_ALARM_alarm_op_2" bit 13
   1272: 'OTEVŘEN BEZPEČNOSTNÍ KRYT (dveře 4)', class Errors, trigger "DB_ALARM_alarm_op_2" bit 11
   1273: 'op_3_alarm_2', class Errors, trigger "DB_ALARM_alarm_op_3" bit 1
   1274: 'OTEVŘEN BEZPEČNOSTNÍ KRYT (dveře 3)', class Errors, trigger "DB_ALARM_alarm_op_2" bit 10
   1275: 'OTEVŘEN BEZPEČNOSTNÍ KRYT (dveře 2)', class Errors, trigger "DB_ALARM_alarm_op_2" bit 9
   1276: 'OTEVŘEN BEZPEČNOSTNÍ KRYT (dveře 1)', class Errors, trigger "DB_ALARM_alarm_op_2" bit 8
   1277: 'op_2_alrm_8', class Errors, trigger "DB_ALARM_alarm_op_2" bit 7
   1278: 'op_2_alrm_6', class Errors, trigger "DB_ALARM_alarm_op_2" bit 5
   1279: 'op_2_alrm_5', class Errors, trigger "DB_ALARM_alarm_op_2" bit 4
   1280: 'PŘERUŠEN BEZPEČNOSTNÍ PAPRSEK V TUNELU', class Errors, trigger "DB_ALARM_alarm_op_2" bit 12
   1281: 'op_3_alarm_3', class Errors, trigger "DB_ALARM_alarm_op_3" bit 2
   1282: 'op_3_alarm_5', class Errors, trigger "DB_ALARM_alarm_op_3" bit 4
   1283: 'PŘEKROČENÍ HLADINY -20B20 ZKONTROLUJTE ZDA NEPROJELI DVĚ TUŽKY NA SOBĚ / ZKŘÍPNUTÍ TUŽKY POD SEGMENTEM !', class Errors, trigger "DB_ALARM_alarm_op_2" bit 3
   1284: 'op_4_alrm_12', class Errors, trigger "DB_ALARM_alarm_op_4" bit 3
   1285: 'op_4_alrm_11', class Errors, trigger "DB_ALARM_alarm_op_4" bit 2
   1286: 'op_4_alrm_10', class Errors, trigger "DB_ALARM_alarm_op_4" bit 1
   1287: 'Odsávací zařízení nereaguje. Otevřete dveře a zkontrolujte jej.', class Errors, trigger "DB_ALARM_alarm_op_4" bit 0
   1288: 'op_4_alrm_15', class Errors, trigger "DB_ALARM_alarm_op_4" bit 6
   1289: 'Odsávací zařízení nereaguje. Otevřete dveře a zkontrolujte jej.', class Errors, trigger "DB_ALARM_alarm_op_4" bit 7
   1290: 'op_3_alarm_16', class Errors, trigger "DB_ALARM_alarm_op_3" bit 15
   1291: 'op_3_alarm_15', class Errors, trigger "DB_ALARM_alarm_op_3" bit 14
   1292: 'op_3_alarm_14', class Errors, trigger "DB_ALARM_alarm_op_3" bit 13
   1293: 'op_3_alarm_13', class Errors, trigger "DB_ALARM_alarm_op_3" bit 12
   1294: 'op_3_alarm_12', class Errors, trigger "DB_ALARM_alarm_op_3" bit 11
   1295: 'op_3_alarm_11', class Errors, trigger "DB_ALARM_alarm_op_3" bit 10
   1296: 'op_3_alarm_10', class Errors, trigger "DB_ALARM_alarm_op_3" bit 9
   1297: 'op_3_alarm_9', class Errors, trigger "DB_ALARM_alarm_op_3" bit 8
   1298: 'op_3_alarm_8', class Errors, trigger "DB_ALARM_alarm_op_3" bit 7
   1299: 'op_3_alarm_7', class Errors, trigger "DB_ALARM_alarm_op_3" bit 6
   1300: 'op_3_alarm_6', class Errors, trigger "DB_ALARM_alarm_op_3" bit 5
   1301: 'op_3_alarm_4', class Errors, trigger "DB_ALARM_alarm_op_3" bit 3
   1302: 'NEDOVŘENÍ PODÉLNÝCH ČELISTÍ -17B2 - (zkontrolujte prostor Čelistí a spusťte výrobu)', class Errors, trigger "DB_ALARM_alarm_op_2" bit 2
   1303: 'SERVO SELHÁNÍ BLOKU OVLÁDÁNÍ "JOG"( KONTAKTUJTE LIFTEC)', class Errors, trigger "DB_ALARM_alarm_op_2" bit 0
   1304: 'op_4_alrm_13', class Errors, trigger "DB_ALARM_alarm_op_4" bit 4
   1305: 'alarm_line_16', class Errors, trigger "DB_ALARM_alarm_line" bit 15
   1306: 'Nedostatečný tlak vzduchu', class Errors, trigger "DB_ALARM_alarm_line" bit 14
   1307: 'alarm_line_14', class Errors, trigger "DB_ALARM_alarm_line" bit 13
   1308: 'alarm_line_13', class Errors, trigger "DB_ALARM_alarm_line" bit 12
   1309: 'alarm_line_12', class Errors, trigger "DB_ALARM_alarm_line" bit 11
   1310: 'alarm_line_11', class Errors, trigger "DB_ALARM_alarm_line" bit 10
   1311: 'APLIKÁTOR ETIKET V PORUŠE ZKONTROLUJTE', class Errors, trigger "DB_ALARM_alarm_line" bit 9
   1312: 'Globální alarm - zařízení nebo část zařízení je v poruše', class Errors, trigger "DB_ALARM_alarm_line" bit 8
   1313: 'alarm_line_8', class Errors, trigger "DB_ALARM_alarm_line" bit 7
   1314: 'Safety I/O potřebuje restart', class Errors, trigger "DB_ALARM_alarm_line" bit 6
   1315: 'alarm_line_6', class Errors, trigger "DB_ALARM_alarm_line" bit 5
   1316: 'alarm_line_5', class Errors, trigger "DB_ALARM_alarm_line" bit 4
   1317: 'alarm_line_4', class Errors, trigger "DB_ALARM_alarm_line" bit 3
   1318: 'alarm_line_3', class Errors, trigger "DB_ALARM_alarm_line" bit 2
   1319: 'alarm_line_2', class Errors, trigger "DB_ALARM_alarm_line" bit 1
   1320: 'op_4_alrm_8', class Errors, trigger "DB_ALARM_alarm_op_4" bit 14
   1321: 'OTEVŘEN BEZPEČNOSTNÍ KRYT (dveře 1)', class Errors, trigger "DB_ALARM_alarm_op_4" bit 15
   1322: 'alarm_line_1', class Errors, trigger "DB_ALARM_alarm_line" bit 0
   1323: 'SERVO - NEZDAŘIL SE RESET N-CODÉRU - PŘEPNĚTE DO MANULÁLU A ZPĚT', class Errors, trigger "DB_ALARM_alarm_op_2" bit 1
   1324: 'op_4_alrm_7', class Errors, trigger "DB_ALARM_alarm_op_4" bit 13
   1325: 'op_1_alrm_1', class Errors, trigger "DB_ALARM_alarm_op_1" bit 0
   1326: 'op_4_alrm_4', class Errors, trigger "DB_ALARM_alarm_op_4" bit 10
   1327: 'op_4_alrm_5', class Errors, trigger "DB_ALARM_alarm_op_4" bit 11
   1328: 'Měření hladiny tužek - senzro je v poruše zkontrolujte / srovnejte hladinu tužek', class Errors, trigger "DB_ALARM_alarm_op_1" bit 15
   1329: 'op_1_alrm_15', class Errors, trigger "DB_ALARM_alarm_op_1" bit 14
   1330: 'op_1_alrm_14', class Errors, trigger "DB_ALARM_alarm_op_1" bit 13
   1331: 'op_1_alrm_13', class Errors, trigger "DB_ALARM_alarm_op_1" bit 12
   1332: 'op_1_alrm_12', class Errors, trigger "DB_ALARM_alarm_op_1" bit 11
   1333: 'op_1_alrm_11', class Errors, trigger "DB_ALARM_alarm_op_1" bit 10
   1334: 'op_1_alrm_10', class Errors, trigger "DB_ALARM_alarm_op_1" bit 9
   1335: 'OTEVŘEN BEZPEČNOSTNÍ KRYT (dveře 1)', class Errors, trigger "DB_ALARM_alarm_op_1" bit 8
   1336: 'op_1_alrm_8', class Errors, trigger "DB_ALARM_alarm_op_1" bit 7
   1337: 'op_1_alrm_7', class Errors, trigger "DB_ALARM_alarm_op_1" bit 6
   1338: 'op_1_alrm_6', class Errors, trigger "DB_ALARM_alarm_op_1" bit 5
   1339: 'op_1_alrm_5', class Errors, trigger "DB_ALARM_alarm_op_1" bit 4
   1340: 'op_1_alrm_4', class Errors, trigger "DB_ALARM_alarm_op_1" bit 3
   1341: 'op_1_alrm_3', class Errors, trigger "DB_ALARM_alarm_op_1" bit 2
   1342: 'op_1_alrm_2', class Errors, trigger "DB_ALARM_alarm_op_1" bit 1
   1343: 'op_4_alrm_6', class Errors, trigger "DB_ALARM_alarm_op_4" bit 12
   1344: 'op_4_alrm_14', class Errors, trigger "DB_ALARM_alarm_op_4" bit 5

text list "error_ropex": 101 'Žádný aktuální signál'; 102 'žádný napěťový signál'; 103 'žádný proud/napěťový signál'; 107 'teplotní krok, dolů'; 108 'teplotní krok, nahoru'; 307 'teplota příliš vysoká / nízká'; 308 'teplota příliš vysoká / nízká'; 309 'teplota příliš vysoká / nízká'; 310 'teplota příliš vysoká / nízká'; 201 'žádná frekvence linky / frekvence linky nekolísá'; 202 'frekvence linky je příliš vysoká / kolísá'; 203 'frekvence linky je příliš nízká / kolísá'; 304 'příliš dlouhá doba zahřívání'; 901 'žádné síťové napětí / synchronizační signál'; 913 'triak vadný'; 914 'vnitřní závada, zařízení vadné'; 915 'vnitřní závada, zařízení vadné'; 916 'vnitřní závada, zařízení vadné'; 917 'můstek pro výstup alarmu je nesprávný'; 918 'můstek pro výstup alarmu je nesprávný'; 0 'OK'

text list "OP_1": 0 'STROJ NESPUŠTĚN'; 1000 'INICIALIZACE - BĚŽÍ'; 1005 'INICIALIZACE - KONTROLA HORNÍ KAMERY'; 1010 'INICIALIZACE - KONTROLA LEVÉ KAMERY'; 1015 'INICIALIZACE - KONTROLA PRAVÉ KAMERY'; 1020 'INICIALIZACE - REZERVA'; 5 'ČEKÁM NA START'; 10 'ZÁSOBNÍK JE NAD MINIMEM'; 15 'VYROVNÁVÁNÍ HLADINY TUŽEK'; 20 'empty'; 25 'empty'; 30 'empty'; 35 'empty'; 40 'empty'; 45 'empty'; 50 'empty'; 55 'empty'; 60 'empty'; 65 'empty'; 70 'empty'; 75 'empty'; 80 'empty'; 85 'empty'; 90 'empty'; 95 'empty'; 100 'empty'; 2 'empty'

text list "OP_2": 0 'STROJ NESPUŠTĚN'; 2 'MANUÁLNÍ REŽIM'; 5 'ČEKÁM NA START'; 10 'CONNECT 192.168.0.100'; 15 'SEND STOP TISKU'; 20 'ČEKÁNÍ NA ODPOVĚĎ'; 25 'DISCONNECT 192.168.0.100'; 30 'CONNECT 192.168.0.100'; 35 'SNED OTEVÍRÁNÍ ZPRÁVY'; 40 'ČEKÁNÍ NA ODPOVĚĎ'; 45 'DISCONNECT 192.168.0.100'; 50 'ROZHODOVÁNÍ ZDA ODESLAT VARIABILNÍ POLE'; 55 'CONNECT 192.168.0.100'; 60 'SEND ODESÍLÁNÍ VARIABILNÍHO POLE'; 65 'ČEKÁNÍ NA ODPOVĚĎ'; 70 'DISCONNECT 192.168.0.100'; 75 'CONNECT 192.168.0.100'; 80 'SEND START TISKU'; 85 'ČEKÁNÍ NA ODPOVĚĎ'; 90 'DISCONNECT 192.168.0.100'; 95 'MAZÁNÍ POŽADAVKŮ'; 100 'REINICIALIZACE'; 1000 'INICIALIZACE - SPOUŠTÍM INICIALIZACI'; 1005 'INICIALIZACE - PŘIPOJOVÁNÍ K 192.168.0.100'; 1010 'INICIALIZACE - KONTROLA SPOJENÍ'; 1015 'INICIALIZACE - ODPOJENÍ OD 192.168.0.100'; 1020 'INICIALIZACE - OK'; 1021 ''

text list "OP_3": 0 'STROJ NESPUŠTĚN'; 2 'MANUÁLNÍ REŽIM'; 5 'ČEKÁM NA POŽADAVEK OP2'; 10 'DOPRAVA'; 15 'ZASTAVUJI ČEKÁM NA LAMELU -21B4'; 20 'empty'; 25 'empty'; 30 'empty'; 35 'empty'; 40 'empty'; 45 'empty'; 50 'empty'; 55 'empty'; 60 'empty'; 65 'empty'; 70 'empty'; 75 'empty'; 80 'empty'; 85 'empty'; 90 'empty'; 95 'empty'; 100 'empty'; 1000 'INICIALIZACE - KONTROLA OVLADAČE MOTORU'; 1005 'INICIALIZACE - HLEDÁM REFERENČNÍ POLOHU -21B4'; 1010 'empty'; 1015 'empty'; 1020 'empty'

text list "STATUS - LINE": 600 'ZAŘÍZENÍ NENÍ PŘIPRAVENO'; 3 'KONTROLA KRYTU 1 / ZAŘÍZENÍ SPUŠTĚNO'; 5 'KONTROLA KRYTU 2 / ZAŘÍZENÍ SPUŠTĚNO'; 10 'KONTROLA KRYTU 3 / ZAŘÍZENÍ SPUŠTĚNO'; 15 'KONTROLA KRYTU 4 / ZAŘÍZENÍ SPUŠTĚNO'; 25 'KONTROLA MOTORŮ / AUTOMATICKÝ REŽIM'; 100 'MANUÁLNÍ REŽIM'; 2000 'SIMULACE'; 20 'KONTROLA HŘÍBKU'; 30 'START INICIALIZACE OP1, OP2, OP3'; 35 'INICIALIZACE OP1'; 40 'INICIALIZACE OP2'; 45 'INICIALIZACE OP3'; 50 'POSLEDNÍ KONTROLA STROJE'; 55 'AUTOMAT'; 60 'empty'; 65 'empty'; 70 'empty'; 75 'empty'; 80 'REŽIM SEŘÍZENÍ'; 85 'empty'; 90 'empty'; 95 'empty'; 105 'empty'; 110 'empty'; 115 'empty'; 120 'empty'; 125 'empty'; 0 'ČEKÁM NA SPUŠTĚNÍ'

graphic list "aut/man": 1 'Graphic_10'; 0 'Graphic_11'

graphic list "safety": 0 'Graphic_19'; 1 'Graphic_20'

graphic list "sen_green": 0 'Graphic_13'; 1 'Graphic_14'

graphic list "sen_green_neg": 1 'Graphic_13'; 0 'Graphic_14'

graphic list "sen_green_red": 0 'Graphic_22'; 1 'Graphic_14'

graphic list "sen_red_jedna_not_activ": 1 'Graphic_13'; 0 'Graphic_22'

graphic list "sen_yelou_jedna_not_activ": 1 'Graphic_13'; 0 'Graphic_23'

graphic list "stop": 1 'Graphic_20'; 0 'Graphic_19'

recipe "Recepty": Zpráva v tiskárně <- "DB_HMI_recype_recipe_Zprava", Program kamery etikety <- "DB_HMI_recype_recipe_PRG_CAM_etiketa"

screen "Root screen" 800x480, template "Template_1"
   on GenerateScreen: SetTag("OP1_DB.Kamera.kontrola_tridirny", 1)
   GraphicView "Graphic view_1" at 2,78 size 703x375; Picture "WhatsApp_Image_2026-07-09_at_09.36.40-removebg-preview"
   GraphicIOField "Graphic I/O field_1" at 504,53 size 30x30; PictureList "sen_green"
      ProcessValue <- "OP1_DB_SENSORS_Pozice_pistu"
   TextField "Text field_2" at 540,57 size 165x23; Text '- BQ5 - Pozice pístu'
   TextField "Text field_3" at 560,365 size 126x42; Text '- BQ4- Pozice Vyřazení'
   TextField "Text field_4" at 534,442 size 137x23; Text '- BQ2 - Kontrola'
   TextField "Text field_5" at 355,423 size 134x23; Text '- BR1 - Enkodér'
   Button "HmiScreenItemData_1" at 0,193 size 111x47; TextOff 'OP_1 DOPRAVA'; TextOn 'D1'; PictureOff "Navigates to D1 for KTP900 Basic+ PN 17.0.0.0"; PictureOn "Navigates to D1 for KTP900 Basic+ PN 17.0.0.0"; Authorization "Operate"
      on Release: ActivateScreen("OP_1_doprava", 0)
   SymbolicIOField "Symbolic I/O field_1" at 0,51 size 431x32; TextOff '0'; TextOn '1'; TextList "OP_1"
      ProcessValue <- "OP1_DB_SQCR"
   SymbolicIOField "Symbolic I/O field_2" at 0,446 size 431x32; TextOff '0'; TextOn '1'; TextList "OP_2"
      ProcessValue <- "OP2_DB_SQCR"
   TextField "Text field_1" at 548,409 size 148x23; Text '- BQ3 - Přechod 2'
   TextField "Text field_6" at 80,346 size 148x23; Text '- BQ1 - Přechod 1'
   IOField "I/O field_1" at 228,418 size 128x32; FormatPattern 9999999999
      ProcessValue <- "HSC_1"
   IOField "I/O field_2" at 5,254 size 172x32; FormatPattern s99999; Unit Plat / Den
      ProcessValue <- "OP1_DB_aktual_kusy"
   GraphicIOField "Graphic I/O field_6" at 210,121 size 30x30; PictureList "sen_green_red"
      ProcessValue <- "CONTROL_LINE_DB_SEN_STRUCT_dvere_L_B"
   TextField "Text field_7" at 41,125 size 128x23; Text '- SQ1 - Dveře L'
   GraphicIOField "Graphic I/O field_7" at 210,155 size 30x30; PictureList "sen_green_red"
      ProcessValue <- "CONTROL_LINE_DB_SEN_STRUCT_dvere_P_B"
   TextField "Text field_8" at 41,159 size 125x23; Text '- SQ2- Dveře P'
   GraphicIOField "Graphic I/O field_8" at 178,121 size 30x30; PictureList "sen_green_red"
      ProcessValue <- "CONTROL_LINE_DB_SEN_STRUCT_dvere_L_A"
   GraphicIOField "Graphic I/O field_9" at 178,155 size 30x30; PictureList "sen_green_red"
      ProcessValue <- "CONTROL_LINE_DB_SEN_STRUCT_dvere_P_A"
   TextField "Text field_9" at 185,82 size 48x20; Text 'KANÁL'
   TextField "Text field_10" at 169,98 size 48x20; Text 'A'
   TextField "Text field_11" at 201,98 size 48x20; Text 'B'

screen "A1" 800x480, template "Template_1"
   on GenerateScreen: SetTag("OP1_DB.Kamera.kontrola_tridirny", 2)
   Button "Back" at 1,41 size 159x47; TextOff 'Back'
      on Release: ActivateScreen("Root screen", 0)
   Button "HmiScreenItemData_1" at 11,135 size 80x47; TextOff 'A11'; PictureOff "Navigates to A11 for KTP900 Basic+ PN 17.0.0.0"; PictureOn "Navigates to A11 for KTP900 Basic+ PN 17.0.0.0"
      on Release: ActivateScreen("A11", 0)
   Button "HmiScreenItemData_2" at 11,194 size 78x47; TextOff 'A12'; PictureOff "Navigates to A12 for KTP900 Basic+ PN 17.0.0.0"; PictureOn "Navigates to A12 for KTP900 Basic+ PN 17.0.0.0"
      on Release: ActivateScreen("A12", 0)
   GraphicView "Graphic view_1" at 279,37 size 266x225; Picture "WhatsApp_Image_2026-07-09_at_09.36.40__1_-removebg-preview"
   GraphicView "Graphic view_2" at 147,60 size 222x198; Picture "WhatsApp_Image_2026-07-09_at_09.36.40__3_-removebg-preview"
   GraphicView "Graphic view_3" at 448,64 size 222x198; Picture "WhatsApp_Image_2026-07-09_at_09.36.40__3_-removebg-preview"
   IOField "I/O field_1" at 287,406 size 277x32; FormatPattern s9999999999; Unit  mm + - 
      ProcessValue <- "DB_HMI_recype_VZDALENOST_KAMERA_ETIKETA_POZADOVANA"

screen "A11" 800x480, template "Template_1"
   on GenerateScreen: SetTag("OP1_DB.Kamera.kontrola_tridirny", 3)
   TextField "HmiScreenItemData" at 75,246 size 595x22; Text 'A11'
   Button "Back" at 1,41 size 159x47; TextOff 'Back'
      on Release: ActivateScreen("A1", 0)

screen "A12" 800x480, template "Template_1"
   on GenerateScreen: SetTag("OP1_DB.Kamera.kontrola_tridirny", 4)
   TextField "HmiScreenItemData" at 75,246 size 595x22; Text 'A12'
   Button "Back" at 1,41 size 159x47; TextOff 'Back'
      on Release: ActivateScreen("A1", 0)

screen "B1" 800x480, template "Template_1"
   on GenerateScreen: SetTag("OP1_DB.Kamera.kontrola_tridirny", 5)
   Button "HmiScreenItemData_1" at 1,108 size 159x47; TextOff 'B11'; PictureOff "Navigates to B11 for KTP900 Basic+ PN 17.0.0.0"; PictureOn "Navigates to B11 for KTP900 Basic+ PN 17.0.0.0"
      on Release: ActivateScreen("B11", 0)
   Button "HmiScreenItemData_2" at 1,171 size 159x47; TextOff 'B12'; PictureOff "Navigates to B12 for KTP900 Basic+ PN 17.0.0.0"; PictureOn "Navigates to B12 for KTP900 Basic+ PN 17.0.0.0"
      on Release: ActivateScreen("B12", 0)
   GraphicView "Graphic view_1" at 398,52 size 244x209; Picture "WhatsApp_Image_2026-07-09_at_09.36.40__2_-removebg-preview"
   GraphicView "Graphic view_2" at 133,52 size 244x209; Picture "WhatsApp Image 2026-07-09 at 09,36,39-Picsart-BackgroundChanger"
   IOField "I/O field_1" at 242,341 size 319x32; FormatPattern s9999999999; Unit mm + -
      ProcessValue <- "DB_HMI_recype_VZDALENOST_KAMERY_FOLIE_POZADOVANA"

screen "B11" 800x480, template "Template_1"
   on GenerateScreen: SetTag("OP1_DB.Kamera.kontrola_tridirny", 6)
   TextField "HmiScreenItemData" at 75,246 size 595x22; Text 'B11'
   Button "Back" at 1,41 size 159x47; TextOff 'Back'
      on Release: ActivateScreen("B1", 0)

screen "B12" 800x480, template "Template_1"
   on GenerateScreen: SetTag("OP1_DB.Kamera.kontrola_tridirny", 7)
   TextField "HmiScreenItemData" at 75,246 size 595x22; Text 'B12'
   Button "Back" at 1,41 size 159x47; TextOff 'Back'
      on Release: ActivateScreen("B1", 0)

screen "C1" 800x480, template "Template_1"
   on GenerateScreen: SetTag("OP1_DB.Kamera.kontrola_tridirny", 8)
   Button "HmiScreenItemData_1" at 7,306 size 159x47; TextOff 'C12'; PictureOff "Navigates to C12 for KTP900 Basic+ PN 17.0.0.0"; PictureOn "Navigates to C12 for KTP900 Basic+ PN 17.0.0.0"
      on Release: ActivateScreen("C12", 0)
   Button "HmiScreenItemData_2" at 7,365 size 159x47; TextOff 'C13'; PictureOff "Navigates to C13 for KTP900 Basic+ PN 17.0.0.0"; PictureOn "Navigates to C13 for KTP900 Basic+ PN 17.0.0.0"
      on Release: ActivateScreen("C13", 0)
   Button "HmiScreenItemData_3" at 7,424 size 159x47; TextOff 'C11'; PictureOff "Navigates to C11 for KTP900 Basic+ PN 17.0.0.0"; PictureOn "Navigates to C11 for KTP900 Basic+ PN 17.0.0.0"
      on Release: ActivateScreen("C11", 0)
   GraphicView "Graphic view_1" at 398,52 size 244x209; Picture "WhatsApp_Image_2026-07-09_at_09.36.40__2_-removebg-preview"
   GraphicView "Graphic view_2" at 133,52 size 244x209; Picture "WhatsApp Image 2026-07-09 at 09,36,39-Picsart-BackgroundChanger"
   IOField "I/O field_1" at 299,353 size 319x32; FormatPattern s9999999999; Unit mm + -
      ProcessValue <- "DB_HMI_recype_VZDALENOST_KAMERY_FOLIE_POZADOVANA"

screen "C12" 800x480, template "Template_1"
   on GenerateScreen: SetTag("OP1_DB.Kamera.kontrola_tridirny", 9)
   TextField "HmiScreenItemData" at 75,246 size 595x22; Text 'C12'
   Button "Back" at 1,41 size 159x47; TextOff 'Back'
      on Release: ActivateScreen("C1", 0)

screen "C13" 800x480, template "Template_1"
   on GenerateScreen: SetTag("OP1_DB.Kamera.kontrola_tridirny", 10)
   TextField "HmiScreenItemData" at 75,246 size 595x22; Text 'C13'
   Button "Back" at 1,41 size 159x47; TextOff 'Back'
      on Release: ActivateScreen("C1", 0)

screen "C11" 800x480, template "Template_1"
   on GenerateScreen: SetTag("OP1_DB.Kamera.kontrola_tridirny", 11)
   TextField "HmiScreenItemData" at 75,246 size 595x22; Text 'C11'
   Button "Back" at 1,41 size 159x47; TextOff 'Back'
      on Release: ActivateScreen("C1", 0)

screen "D1" 800x480, template "Template_1"
   on GenerateScreen: SetTag("OP1_DB.Kamera.kontrola_tridirny", 12)
   Button "Back" at 1,41 size 159x47; TextOff 'Back'
      on Release: ActivateScreen("Root screen", 0)
   Button "HmiScreenItemData_1" at 36,135 size 159x47; TextOff 'D11'; PictureOff "Navigates to D11 for KTP900 Basic+ PN 17.0.0.0"; PictureOn "Navigates to D11 for KTP900 Basic+ PN 17.0.0.0"
      on Release: ActivateScreen("D11", 0)
   Button "HmiScreenItemData_2" at 36,194 size 159x47; TextOff 'D12'; PictureOff "Navigates to D12 for KTP900 Basic+ PN 17.0.0.0"; PictureOn "Navigates to D12 for KTP900 Basic+ PN 17.0.0.0"
      on Release: ActivateScreen("D12", 0)
   GraphicView "Graphic view_2" at 251,43 size 200x238; Picture "WhatsApp Image 2026-07-09 at 09,43,15-Picsart-BackgroundChanger"

screen "D11" 800x480, template "Template_1"
   on GenerateScreen: SetTag("OP1_DB.Kamera.kontrola_tridirny", 13)
   TextField "HmiScreenItemData" at 75,246 size 595x22; Text 'D11'
   Button "Back" at 1,41 size 159x47; TextOff 'Back'
      on Release: ActivateScreen("D1", 0)

screen "D12" 800x480, template "Template_1"
   on GenerateScreen: SetTag("OP1_DB.Kamera.kontrola_tridirny", 14)
   TextField "HmiScreenItemData" at 75,246 size 595x22; Text 'D12'
   Button "Back" at 1,41 size 159x47; TextOff 'Back'
      on Release: ActivateScreen("D1", 0)

screen "E1" 800x480, template "Template_1"
   on GenerateScreen: SetTag("OP1_DB.Kamera.kontrola_tridirny", 15)
   RecipeView "Recipe view_1" at 1,50 size 725x372; Recipe "Recepty"
   IOField "I/O field_1" at 4,429 size 171x42; FormatPattern ????????????????????
      ProcessValue <- "DB_HMI_recype_recipe_pole_string_1"
   Button "Button_1" at 520,429 size 203x42; TextOff 'Odeslání dat do tiskárny'
      on Click: SetBit("DB_HMI_recype_ODESLI_dATA")
      Appearance <- "DB_HMI_recype_ODESLI_dATA"
   TextField "Text field_1" at 184,436 size 64x27; Text 'Pole 1'
   IOField "I/O field_2" at 257,429 size 171x42; FormatPattern ??????????
      ProcessValue <- "DB_HMI_recype_recipe_pole_string_2"
   TextField "Text field_2" at 438,436 size 64x27; Text 'Pole 2'
   Button "Button_2" at 259,341 size 138x33; TextOff 'Kontrola třídírny'
      on Click: InvertBit("OP1_DB.Kamera.kontrola_tridirny")
      Appearance <- "OP1_DB.Kamera.kontrola_tridirny"

screen "E11" 800x480, template "Template_1"
   on GenerateScreen: SetTag("OP1_DB.Kamera.kontrola_tridirny", 16)
   TextField "HmiScreenItemData" at 75,246 size 595x22; Text 'E11'
   Button "Back" at 1,41 size 159x47; TextOff 'Back'
      on Release: ActivateScreen("E1", 0)

screen "E12" 800x480, template "Template_1"
   on GenerateScreen: SetTag("OP1_DB.Kamera.kontrola_tridirny", 17)
   TextField "HmiScreenItemData" at 75,246 size 595x22; Text 'E12'
   Button "Back" at 1,41 size 159x47; TextOff 'Back'
      on Release: ActivateScreen("E1", 0)

screen "F1" 800x480, template "Template_1"
   on GenerateScreen: SetTag("OP1_DB.Kamera.kontrola_tridirny", 18)
   TextField "HmiScreenItemData" at 75,246 size 595x22; Text 'F1'
   Button "Back" at 1,41 size 159x47; TextOff 'Back'
      on Release: ActivateScreen("Root screen", 0)
   Button "HmiScreenItemData_1" at 36,135 size 159x47; TextOff 'F11'; PictureOff "Navigates to F11 for KTP900 Basic+ PN 17.0.0.0"; PictureOn "Navigates to F11 for KTP900 Basic+ PN 17.0.0.0"
      on Release: ActivateScreen("F11", 0)

screen "F11" 800x480, template "Template_1"
   on GenerateScreen: SetTag("OP1_DB.Kamera.kontrola_tridirny", 19)
   TextField "HmiScreenItemData" at 75,246 size 595x22; Text 'F11'
   Button "Back" at 1,41 size 159x47; TextOff 'Back'
      on Release: ActivateScreen("F1", 0)

screen "System screens" 800x480, template "Template_1"
   on GenerateScreen: SetTag("OP1_DB.Kamera.kontrola_tridirny", 20)
   Button "Back" at 1,41 size 159x47; TextOff 'Back'
      on Release: ActivateScreen("Root screen", 0)
   Button "HmiScreenItemData" at 36,135 size 159x47; TextOff 'SIMATIC PLC system diagnos...'; PictureOff "Navigates to SIMATIC PLC system diagnostics for KTP900 Basic+ PN 17.0.0.0"; PictureOn "Navigates to SIMATIC PLC system diagnostics for KTP900 Basic+ PN 17.0.0.0"
      on Release: ActivateScreen("SIMATIC PLC system diagnostics", 0)
   Button "HmiScreenItemData_1" at 36,194 size 159x47; TextOff 'Project information'; PictureOff "Navigates to Project information for KTP900 Basic+ PN 17.0.0.0"; PictureOn "Navigates to Project information for KTP900 Basic+ PN 17.0.0.0"
      on Release: ActivateScreen("Project information", 0)
   Button "HmiScreenItemData_2" at 36,253 size 159x47; TextOff 'User administration'; PictureOff "Navigates to User administration for KTP900 Basic+ PN 17.0.0.0"; PictureOn "Navigates to User administration for KTP900 Basic+ PN 17.0.0.0"
      on Release: ActivateScreen("User administration", 0)
   Button "HmiScreenItemData_3" at 36,312 size 159x47; TextOff 'System information'; PictureOff "Navigates to System information for KTP900 Basic+ PN 17.0.0.0"; PictureOn "Navigates to System information for KTP900 Basic+ PN 17.0.0.0"
      on Release: ActivateScreen("System information", 0)
   Button "HmiScreenItemData_4" at 36,371 size 159x47; TextOff 'Different jobs'; PictureOff "Navigates to Different jobs for KTP900 Basic+ PN 17.0.0.0"; PictureOn "Navigates to Different jobs for KTP900 Basic+ PN 17.0.0.0"
      on Release: ActivateScreen("Different jobs", 0)

screen "SIMATIC PLC system diagnostics" 800x480, template "Template_1"
   on GenerateScreen: SetTag("OP1_DB.Kamera.kontrola_tridirny", 21)
   SysDiagControl "HmiScreenItemData" at 1,89 size 740x383
   Button "Back" at 1,41 size 159x47; TextOff 'Back'
      on Release: ActivateScreen("System screens", 0)

screen "Project information" 800x480, template "Template_1"
   on GenerateScreen: SetTag("OP1_DB.Kamera.kontrola_tridirny", 22)
   TextField "HmiScreenItemData" at 35,91 size 171x28; Text 'Project name:'
   TextField "HmiScreenItemData_1" at 241,91 size 468x28; Text 'Ceska_vejce_2026_06_25'
   TextField "HmiScreenItemData_2" at 35,121 size 171x28; Text 'Created on:'
   TextField "HmiScreenItemData_3" at 241,121 size 468x28; Text '6/25/2026 1:40:25 PM'
   TextField "HmiScreenItemData_4" at 35,151 size 171x28; Text 'Author:'
   TextField "HmiScreenItemData_5" at 241,151 size 468x28; Text 'pavel.svitak'
   TextField "HmiScreenItemData_6" at 35,181 size 171x28; Text 'Description:'
   TextField "HmiScreenItemData_7" at 241,181 size 468x28; Text '(not configured)'
   Button "Back" at 1,41 size 159x47; TextOff 'Back'
      on Release: ActivateScreen("System screens", 0)

screen "User administration" 800x480, template "Template_1"
   on GenerateScreen: SetTag("OP1_DB.Kamera.kontrola_tridirny", 23)
   UserView "HmiScreenItemData" at 1,89 size 740x383
   Button "Back" at 1,41 size 159x47; TextOff 'Back'
      on Release: ActivateScreen("System screens", 0)

screen "System information" 800x480, template "Template_1"
   on GenerateScreen: SetTag("OP1_DB.Kamera.kontrola_tridirny", 24)
   TextField "HmiScreenItemData" at 35,91 size 171x28; Text 'HMI device type:'
   TextField "HmiScreenItemData_1" at 241,91 size 468x28; Text 'KTP900 Basic+ PN 17.0.0.0'
   TextField "HmiScreenItemData_2" at 35,121 size 171x28; Text 'Connection:'
   TextField "HmiScreenItemData_3" at 241,121 size 468x28; Text 'PROFINET (X1)'
   TextField "HmiScreenItemData_4" at 35,151 size 171x28; Text 'PLC:'
   TextField "HmiScreenItemData_5" at 241,151 size 468x28; Text 'SIMATIC S7 1200'
   Button "Back" at 1,41 size 159x47; TextOff 'Back'
      on Release: ActivateScreen("System screens", 0)

screen "Different jobs" 800x480, template "Template_1"
   on GenerateScreen: SetTag("OP1_DB.Kamera.kontrola_tridirny", 25)
   Button "Online" at 36,135 size 159x47; TextOff 'Online'
      on Release: function_bb44b551(0)
   Button "Offline" at 36,194 size 159x47; TextOff 'Offline'
      on Release: function_bb44b551(1)
   Button "Transfer" at 36,253 size 159x47; TextOff 'Transfer'
      on Release: function_bb44b551(2)
   Button "Toggle language" at 36,312 size 159x47; TextOff 'Toggle language'
      on Release: function_fb9197e8(-1)
   Button "Stop Runtime" at 36,371 size 159x47; TextOff 'Stop Runtime'
      on Release: StopRuntime(0)
   Button "Back" at 1,41 size 159x47; TextOff 'Back'
      on Release: ActivateScreen("System screens", 0)

Template "Template_1" 800x480
   Button "Start screen" at 727,52 size 71x50; TextOff 'Start screen'; PictureOn "NavigateHome_KTP700_Basic_PN_TR"; PictureOff "Graphic_2"
      on Release: ActivateScreen("Root screen", 0)
   Button "Alarms" at 727,106 size 71x50; TextOff 'Alarms'; PictureOff "Graphic_3"; PictureOn "Graphic_3"
      on Release: function_ef3f5d25("Alarm window_Unacknowledged", -1)
      Appearance <- "CONTROL_LINE_DB_HMI_ALARM"
   Button "Log on" at 727,159 size 71x50; TextOff 'Log on'; PictureOn "Login_KTP700_Basic_PN_TR"; PictureOff "Graphic_4"; Authorization "Operate"
      on Release: function_a2a04561()
   Button "Language" at 727,213 size 71x50; TextOff 'Language'; PictureOn "ToggleLanguage_KTP700_Basic_PN_TR"; PictureOff "Graphic_5"; Authorization "User administration"
      on Release: function_fb9197e8(-1)
   Button "Template_Button" at 727,267 size 71x50; TextOff 'Text'; PictureOff "Graphic_12"; Authorization "User administration"
      on Release: ActivateScreen("System screens", 0)
   Button "Template_Button_1" at 727,321 size 71x50; TextOff 'Text'; PictureOff "Graphic_9"; Authorization "Operate"
      on Release: ActivateScreen("E1", 0)
      Visibility <- "OP2_DB_TRIG_inicial_ok_op"
   Button "Template_Button_2" at 727,374 size 71x50; TextOff 'Text'; PictureOff "Graphic_8"
      on Release: function_efd93a16()
   Button "Exit" at 727,428 size 71x50; TextOff 'Exit'; PictureOn "ExitRuntime_KTP700_Basic_PN_TR"; PictureOff "Graphic_6"; Authorization "User administration"
      on Release: StopRuntime(0)
   DateTimeField "HmiScreenItemData" at 695,25 size 105x25
   DateTimeField "HmiScreenItemData_1" at 695,0 size 105x25
   GraphicIOField "Template_Graphic I/O field_1" at 661,5 size 40x40; PictureList "aut/man"
      ProcessValue <- "AUT_MAN_HMI"
   GraphicView "Template_Graphic view_1" at 0,0 size 50x50; Picture "images"
   SymbolicIOField "Template_Symbolic I/O field_1" at 161,9 size 498x32; TextOff '0'; TextOn '1'; TextList "STATUS - LINE"
      Appearance <- "CONTROL_LINE_DB_SQCR"
      ProcessValue <- "CONTROL_LINE_DB_SQCR"

screen "OP_1_doprava" 800x480, template "Template_1"
   GraphicView "Graphic view_1" at 1,98 size 703x375; Picture "WhatsApp_Image_2026-07-09_at_09.36.40-removebg-preview"
   Button "HmiScreenItemData" at 1,295 size 129x47; TextOff 'kamera horní'; TextOn 'A1'; PictureOff "Navigates to A1 for KTP900 Basic+ PN 17.0.0.0"; PictureOn "Navigates to A1 for KTP900 Basic+ PN 17.0.0.0"; Authorization "User administration"
      on Release: ActivateScreen("A1", 0)
   Button "HmiScreenItemData_1" at 0,403 size 134x47; TextOff 'kamera pravá'; TextOn 'B1'; PictureOff "Navigates to B1 for KTP900 Basic+ PN 17.0.0.0"; PictureOn "Navigates to B1 for KTP900 Basic+ PN 17.0.0.0"; Authorization "User administration"
      on Release: ActivateScreen("B1", 0)
   Button "HmiScreenItemData_2" at 1,348 size 129x47; TextOff 'kamera levá'; TextOn 'C1'; PictureOff "Navigates to C1 for KTP900 Basic+ PN 17.0.0.0"; PictureOn "Navigates to C1 for KTP900 Basic+ PN 17.0.0.0"; Authorization "User administration"
      on Release: ActivateScreen("C1", 0)
   IOField "I/O field_1" at 329,53 size 295x25; FormatPattern ????????????????????????????????????????????????????????????????????????????????
      ProcessValue <- "DB_HMI_recype_fronta{1}_prenaseny_text"
      Visibility <- "DB_HMI_recype_obsazenost_fronty"
      Appearance <- "DB_HMI_recype_fronta{1}_vyrazeni"
   IOField "I/O field_2" at 626,53 size 69x25; FormatPattern 99999
      ProcessValue <- "DB_HMI_recype_fronta{1}_balik_den"
      Visibility <- "DB_HMI_recype_obsazenost_fronty"
      Appearance <- "DB_HMI_recype_fronta{1}_vyrazeni"
   IOField "I/O field_3" at 697,53 size 27x25; FormatPattern 1
      ProcessValue <- "DB_HMI_recype_fronta{1}_vyrazeni"
      Visibility <- "DB_HMI_recype_obsazenost_fronty"
      Appearance <- "DB_HMI_recype_fronta{1}_vyrazeni"
   Line "Line_4" at 555,82 size 159x148
      Visibility <- "DB_HMI_recype_obsazenost_fronty"
   IOField "I/O field_4" at 294,80 size 295x24; FormatPattern ????????????????????????????????????????????????????????????????????????????????
      ProcessValue <- "DB_HMI_recype_fronta{2}_prenaseny_text"
      Visibility <- "DB_HMI_recype_obsazenost_fronty"
      Appearance <- "DB_HMI_recype_fronta{2}_vyrazeni"
   IOField "I/O field_5" at 591,80 size 69x25; FormatPattern 99999
      ProcessValue <- "DB_HMI_recype_fronta{2}_balik_den"
      Visibility <- "DB_HMI_recype_obsazenost_fronty"
      Appearance <- "DB_HMI_recype_fronta{2}_vyrazeni"
   IOField "I/O field_6" at 662,80 size 27x25; FormatPattern 1
      ProcessValue <- "DB_HMI_recype_fronta{2}_vyrazeni"
      Visibility <- "DB_HMI_recype_obsazenost_fronty"
      Appearance <- "DB_HMI_recype_fronta{2}_vyrazeni"
   IOField "I/O field_7" at 263,106 size 295x25; FormatPattern ????????????????????????????????????????????????????????????????????????????????
      ProcessValue <- "DB_HMI_recype_fronta{3}_prenaseny_text"
      Visibility <- "DB_HMI_recype_obsazenost_fronty"
      Appearance <- "DB_HMI_recype_fronta{3}_vyrazeni"
   IOField "I/O field_8" at 560,106 size 69x25; FormatPattern 99999
      ProcessValue <- "DB_HMI_recype_fronta{3}_balik_den"
      Visibility <- "DB_HMI_recype_obsazenost_fronty"
      Appearance <- "DB_HMI_recype_fronta{3}_vyrazeni"
   IOField "I/O field_9" at 631,106 size 27x25; FormatPattern 1
      ProcessValue <- "DB_HMI_recype_fronta{3}_vyrazeni"
      Visibility <- "DB_HMI_recype_obsazenost_fronty"
      Appearance <- "DB_HMI_recype_fronta{3}_vyrazeni"
   IOField "I/O field_10" at 235,133 size 295x25; FormatPattern ????????????????????????????????????????????????????????????????????????????????
      ProcessValue <- "DB_HMI_recype_fronta{4}_prenaseny_text"
      Visibility <- "DB_HMI_recype_obsazenost_fronty"
      Appearance <- "DB_HMI_recype_fronta{4}_vyrazeni"
   IOField "I/O field_11" at 532,133 size 69x25; FormatPattern 99999
      ProcessValue <- "DB_HMI_recype_fronta{4}_balik_den"
      Visibility <- "DB_HMI_recype_obsazenost_fronty"
      Appearance <- "DB_HMI_recype_fronta{4}_vyrazeni"
   IOField "I/O field_12" at 602,133 size 27x25; FormatPattern 1
      ProcessValue <- "DB_HMI_recype_fronta{4}_vyrazeni"
      Visibility <- "DB_HMI_recype_obsazenost_fronty"
      Appearance <- "DB_HMI_recype_fronta{4}_vyrazeni"
   IOField "I/O field_13" at 205,160 size 295x25; FormatPattern ????????????????????????????????????????????????????????????????????????????????
      ProcessValue <- "DB_HMI_recype_fronta{5}_prenaseny_text"
      Visibility <- "DB_HMI_recype_obsazenost_fronty"
      Appearance <- "DB_HMI_recype_fronta{5}_vyrazeni"
   IOField "I/O field_14" at 503,160 size 69x25; FormatPattern 99999
      ProcessValue <- "DB_HMI_recype_fronta{5}_balik_den"
      Visibility <- "DB_HMI_recype_obsazenost_fronty"
      Appearance <- "DB_HMI_recype_fronta{5}_vyrazeni"
   IOField "I/O field_15" at 574,160 size 27x25; FormatPattern 1
      ProcessValue <- "DB_HMI_recype_fronta{5}_vyrazeni"
      Visibility <- "DB_HMI_recype_obsazenost_fronty"
      Appearance <- "DB_HMI_recype_fronta{5}_vyrazeni"
   Line "Line_5" at 385,234 size 160x17
      Visibility <- "DB_HMI_recype_obsazenost_fronty"
   Line "Line_6" at 129,65 size 173x2
      Visibility <- "DB_HMI_recype_obsazenost_fronty"
   TextField "Text field_1" at 307,56 size 17x20; Text '1.'
      Visibility <- "DB_HMI_recype_obsazenost_fronty"
   TextField "Text field_2" at 274,82 size 17x20; Text '2.'
      Visibility <- "DB_HMI_recype_obsazenost_fronty"
   TextField "Text field_3" at 243,109 size 17x20; Text '3.'
      Visibility <- "DB_HMI_recype_obsazenost_fronty"
   TextField "Text field_4" at 215,136 size 17x20; Text '4.'
      Visibility <- "DB_HMI_recype_obsazenost_fronty"
   TextField "Text field_5" at 184,163 size 17x20; Text '5.'
      Visibility <- "DB_HMI_recype_obsazenost_fronty"
   Line "Line_7" at 127,70 size 144x22
      Visibility <- "DB_HMI_recype_obsazenost_fronty"
   Line "Line_8" at 133,80 size 105x36
      Visibility <- "DB_HMI_recype_obsazenost_fronty"
   Line "Line_9" at 133,91 size 80x50
      Visibility <- "DB_HMI_recype_obsazenost_fronty"
   Line "Line_10" at 132,101 size 52x72
      Visibility <- "DB_HMI_recype_obsazenost_fronty"
   Button "Button_1" at 12,58 size 129x55; TextOff 'Smazání bafru'
      Visibility <- "DB_HMI_recype_obsazenost_fronty"
      on Press: SetBit("OP1_DB_HMI_hmi_5")
   IOField "I/O field_16" at 29,116 size 96x32; FormatPattern 9
      ProcessValue <- "DB_HMI_recype_obsazenost_fronty"
      Visibility <- "DB_HMI_recype_obsazenost_fronty"

screen "OP_2_tiskárna" 800x480, template "Template_1"
   Button "HmiScreenItemData_3" at 29,67 size 111x47; TextOff 'tiskárna'; TextOn 'D1'; PictureOff "Navigates to D1 for KTP900 Basic+ PN 17.0.0.0"; PictureOn "Navigates to D1 for KTP900 Basic+ PN 17.0.0.0"
      on Release: ActivateScreen("D1", 0)
*)